    PROC Path_RobotLab(PERS wobjdata WO_Pastel)
        Path_vacio_ejecucion p_vacio_labSIR, 1, WO_Pastel, FALSE;
        index_vacio_destino:=25;
        Path_contacto_ejecucion p_contacto_labSIR, 1, 3, WO_Pastel, FALSE;
        Mover_en_contacto;
        TriggC p_contacto_labSIR{4},p_contacto_labSIR{5},Vel_Proceso,triggContactoCir,Z_Proceso,Prototipo_JSDaleman\WObj:=WO_Pastel;
        TriggL p_contacto_labSIR{6},Vel_Proceso,triggContacto,Z_Proceso,Prototipo_JSDaleman\WObj:=WO_Pastel;
        TriggC p_contacto_labSIR{7},p_contacto_labSIR{8},Vel_Proceso,triggContactoCir,Z_Proceso,Prototipo_JSDaleman\WObj:=WO_Pastel;
        Path_contacto_ejecucion p_contacto_labSIR, 9, 25, WO_Pastel, TRUE;
        Path_vacio_ejecucion p_vacio_labSIR, 2, WO_Pastel, FALSE;
        Path_contacto_ejecucion p_contacto_labSIR, 26, 94, WO_Pastel, TRUE;
        Path_vacio_ejecucion p_vacio_labSIR, 3, WO_Pastel, FALSE;
        Path_contacto_ejecucion p_contacto_labSIR, 95, 111, WO_Pastel, TRUE;
        Path_vacio_ejecucion p_vacio_labSIR, 4, WO_Pastel, FALSE;
        Path_contacto_ejecucion p_contacto_labSIR, 112, 125, WO_Pastel, TRUE;
        Path_vacio_ejecucion p_vacio_labSIR, 5, WO_Pastel, FALSE;
        index_vacio_destino:=131;
        Mover_a_contacto;
        TriggL p_contacto_labSIR{126},Vel_Acercamiento,triggContacto,Z_Acercamiento,Prototipo_JSDaleman\WObj:=WO_Pastel;
        Mover_en_contacto;
        TriggC p_contacto_labSIR{127},p_contacto_labSIR{128},Vel_Proceso,triggContactoCir,Z_Proceso,Prototipo_JSDaleman\WObj:=WO_Pastel;
        TriggC p_contacto_labSIR{129},p_contacto_labSIR{130},Vel_Proceso,triggContactoCir,Z_Proceso,Prototipo_JSDaleman\WObj:=WO_Pastel;
        Mover_a_vacio;
        TriggL p_contacto_labSIR{131},Vel_Acercamiento,triggContacto,Z_Acercamiento,Prototipo_JSDaleman\WObj:=WO_Pastel;
        Path_vacio_ejecucion p_vacio_labSIR, 6, WO_Pastel, FALSE;
        index_vacio_destino:=137;
        Mover_a_contacto;
        TriggL p_contacto_labSIR{132},Vel_Acercamiento,triggContacto,Z_Acercamiento,Prototipo_JSDaleman\WObj:=WO_Pastel;
        Mover_en_contacto;
        TriggC p_contacto_labSIR{133},p_contacto_labSIR{134},Vel_Proceso,triggContactoCir,Z_Proceso,Prototipo_JSDaleman\WObj:=WO_Pastel;
        TriggC p_contacto_labSIR{135},p_contacto_labSIR{136},Vel_Proceso,triggContactoCir,Z_Proceso,Prototipo_JSDaleman\WObj:=WO_Pastel;
        Mover_a_vacio;
        TriggL p_contacto_labSIR{137},Vel_Acercamiento,triggContacto,Z_Acercamiento,Prototipo_JSDaleman\WObj:=WO_Pastel;
        Path_vacio_ejecucion p_vacio_labSIR, 7, WO_Pastel, FALSE;
        index_vacio_destino:=143;
        Mover_a_contacto;
        TriggL p_contacto_labSIR{138},Vel_Acercamiento,triggContacto,Z_Acercamiento,Prototipo_JSDaleman\WObj:=WO_Pastel;
        Mover_en_contacto;
        TriggC p_contacto_labSIR{139},p_contacto_labSIR{140},Vel_Proceso,triggContactoCir,Z_Proceso,Prototipo_JSDaleman\WObj:=WO_Pastel;
        TriggC p_contacto_labSIR{141},p_contacto_labSIR{142},Vel_Proceso,triggContactoCir,Z_Proceso,Prototipo_JSDaleman\WObj:=WO_Pastel;
        Mover_a_vacio;
        TriggL p_contacto_labSIR{143},Vel_Acercamiento,triggContacto,Z_Acercamiento,Prototipo_JSDaleman\WObj:=WO_Pastel;
        Path_vacio_ejecucion p_vacio_labSIR, 8, WO_Pastel, FALSE;
        index_vacio_destino:=149;
        Mover_a_contacto;
        TriggL p_contacto_labSIR{144},Vel_Acercamiento,triggContacto,Z_Acercamiento,Prototipo_JSDaleman\WObj:=WO_Pastel;
        Mover_en_contacto;
        TriggC p_contacto_labSIR{145},p_contacto_labSIR{146},Vel_Proceso,triggContactoCir,Z_Proceso,Prototipo_JSDaleman\WObj:=WO_Pastel;
        TriggC p_contacto_labSIR{147},p_contacto_labSIR{148},Vel_Proceso,triggContactoCir,Z_Proceso,Prototipo_JSDaleman\WObj:=WO_Pastel;
        Mover_a_vacio;
        TriggL p_contacto_labSIR{149},Vel_Acercamiento,triggContacto,Z_Acercamiento,Prototipo_JSDaleman\WObj:=WO_Pastel;
        Path_vacio_ejecucion p_vacio_labSIR, 9, WO_Pastel, FALSE;
        index_vacio_destino:=155;
        Mover_a_contacto;
        TriggL p_contacto_labSIR{150},Vel_Acercamiento,triggContacto,Z_Acercamiento,Prototipo_JSDaleman\WObj:=WO_Pastel;
        Mover_en_contacto;
        TriggC p_contacto_labSIR{151},p_contacto_labSIR{152},Vel_Proceso,triggContactoCir,Z_Proceso,Prototipo_JSDaleman\WObj:=WO_Pastel;
        TriggC p_contacto_labSIR{153},p_contacto_labSIR{154},Vel_Proceso,triggContactoCir,Z_Proceso,Prototipo_JSDaleman\WObj:=WO_Pastel;
        Mover_a_vacio;
        TriggL p_contacto_labSIR{155},Vel_Acercamiento,triggContacto,Z_Acercamiento,Prototipo_JSDaleman\WObj:=WO_Pastel;
        Path_vacio_ejecucion p_vacio_labSIR, 10, WO_Pastel, FALSE;
        index_vacio_destino:=161;
        Mover_a_contacto;
        TriggL p_contacto_labSIR{156},Vel_Acercamiento,triggContacto,Z_Acercamiento,Prototipo_JSDaleman\WObj:=WO_Pastel;
        Mover_en_contacto;
        TriggC p_contacto_labSIR{157},p_contacto_labSIR{158},Vel_Proceso,triggContactoCir,Z_Proceso,Prototipo_JSDaleman\WObj:=WO_Pastel;
        TriggC p_contacto_labSIR{159},p_contacto_labSIR{160},Vel_Proceso,triggContactoCir,Z_Proceso,Prototipo_JSDaleman\WObj:=WO_Pastel;
        Mover_a_vacio;
        TriggL p_contacto_labSIR{161},Vel_Proceso,triggContacto,Z_Proceso,Prototipo_JSDaleman\WObj:=WO_Pastel;
    ENDPROC
    PROC Path_Tapa_LabSIR(PERS wobjdata WO_Pastel)
        Mover_en_vacio;
        MoveJ Target_Home_10,Vel_Vacio_Rap,Z_Vacio_Rap,Prototipo_JSDaleman\WObj:=wobj0;
        ReiniciarIndices;
        path_contacto_actual:="p_contacto_labSIR";
        path_vacio_actual:="p_vacio_labSIR";
        Path_RobotLab WO_Pastel;
        Path_LabSIR WO_Pastel;
        Mover_en_vacio;
        MoveJ Target_Home_10,Vel_Vacio_Rap,Z_Vacio_Rap,Prototipo_JSDaleman\WObj:=wobj0;
    ENDPROC
    PROC Path_LabSIR(PERS wobjdata WO_Pastel)
        Path_vacio_ejecucion p_vacio_labSIR, 11, WO_Pastel, FALSE;
        Path_contacto_ejecucion p_contacto_labSIR, 162, 170, WO_Pastel, TRUE;
        Path_vacio_ejecucion p_vacio_labSIR, 12, WO_Pastel, FALSE;
        Path_contacto_ejecucion p_contacto_labSIR, 171, 182, WO_Pastel, TRUE;
        Path_vacio_ejecucion p_vacio_labSIR, 13, WO_Pastel, FALSE;
        Path_contacto_ejecucion p_contacto_labSIR, 183, 188, WO_Pastel, TRUE;
        Path_vacio_ejecucion p_vacio_labSIR, 14, WO_Pastel, FALSE;
        Path_contacto_ejecucion p_contacto_labSIR, 189, 199, WO_Pastel, TRUE;
        Path_vacio_ejecucion p_vacio_labSIR, 15, WO_Pastel, FALSE;
        Path_contacto_ejecucion p_contacto_labSIR, 200, 205, WO_Pastel, TRUE;
        Path_vacio_ejecucion p_vacio_labSIR, 16, WO_Pastel, FALSE;
        Path_contacto_ejecucion p_contacto_labSIR, 206, 219, WO_Pastel, TRUE;
        Path_vacio_ejecucion p_vacio_labSIR, 17, WO_Pastel, FALSE;
        Path_contacto_ejecucion p_contacto_labSIR, 220, 226, WO_Pastel, TRUE;
        Path_vacio_ejecucion p_vacio_labSIR, 18, WO_Pastel, FALSE;
        Path_contacto_ejecucion p_contacto_labSIR, 227, 232, WO_Pastel, TRUE;
        Path_vacio_ejecucion p_vacio_labSIR, 19, WO_Pastel, FALSE;
        Path_contacto_ejecucion p_contacto_labSIR, 233, 256, WO_Pastel, TRUE;
    ENDPROC
    PROC Path_Frente_LabSIR(PERS wobjdata WO_Pastel)
        Mover_en_vacio;
        MoveJ Target_Home_10,Vel_Vacio_Rap,Z_Vacio_Rap,Prototipo_JSDaleman\WObj:=wobj0;
        MoveJ Target_Frente_10,Vel_Vacio,Z_VacioMov,Prototipo_JSDaleman\WObj:=WO_Pastel;
        MoveJ Target_Frente_20,Vel_Vacio,Z_VacioMov,Prototipo_JSDaleman\WObj:=WO_Pastel;
        ReiniciarIndices;
        path_contacto_actual:="p_contacto_labSIR_FrenteL";
        path_vacio_actual:="p_vacio_labSIR_FrenteL";
        Path_Chip WO_Pastel;
        Path_LetreroFrontal1_LabSIR WO_Pastel;
        Path_LetreroFrontal2_LabSIR WO_Pastel;
        Mover_en_vacio;
        MoveJ Target_Frente_20,Vel_Vacio,Z_VacioMov,Prototipo_JSDaleman\WObj:=WO_Pastel;
        MoveJ Target_Frente_10,Vel_Vacio,Z_VacioMov,Prototipo_JSDaleman\WObj:=WO_Pastel;
        MoveJ Target_Home_10,Vel_Vacio_Rap,Z_Vacio_Rap,Prototipo_JSDaleman\WObj:=wobj0;
        MoveJ Target_Frente_30,Vel_Vacio_Rap,Z_Vacio_Rap,Prototipo_JSDaleman\WObj:=WO_Pastel;
        MoveJ Target_Frente_40,Vel_Vacio_Rap,Z_Vacio_Rap,Prototipo_JSDaleman\WObj:=WO_Pastel;
        ReiniciarIndices;
        path_contacto_actual:="p_contacto_labSIR_FrenteR";
        path_vacio_actual:="p_vacio_labSIR_FrenteR";
        Path_Engranaje WO_Pastel;
        Path_LetreroFrontal3_LabSIR WO_Pastel;
        Path_LetreroFrontal4_LabSIR WO_Pastel;
        Mover_en_vacio;
        MoveJ Target_Frente_40,Vel_Vacio_Rap,Z_Vacio_Rap,Prototipo_JSDaleman\WObj:=WO_Pastel;
        MoveJ Target_Frente_30,Vel_Vacio_Rap,Z_Vacio_Rap,Prototipo_JSDaleman\WObj:=WO_Pastel;
        MoveJ Target_Home_10,Vel_Vacio_Rap,Z_Vacio_Rap,Prototipo_JSDaleman\WObj:=wobj0;
    ENDPROC
    PROC Path_Chip(PERS wobjdata WO_Pastel)
        Path_vacio_ejecucion p_vacio_labSIR_FrenteL, 1, WO_Pastel, FALSE;
        Path_contacto_ejecucion p_contacto_labSIR_FrenteL, 1, 50, WO_Pastel, TRUE;
        Path_vacio_ejecucion p_vacio_labSIR_FrenteL, 1, WO_Pastel, FALSE;
        Path_contacto_ejecucion p_contacto_labSIR_FrenteL, 51, 56, WO_Pastel, TRUE;
    ENDPROC
    PROC Path_LetreroFrontal1_LabSIR(PERS wobjdata WO_Pastel)
        Path_vacio_ejecucion p_vacio_labSIR_FrenteL, 3, WO_Pastel, FALSE;
        Path_contacto_ejecucion p_contacto_labSIR_FrenteL, 57, 60, WO_Pastel, TRUE;
        Path_vacio_ejecucion p_vacio_labSIR_FrenteL, 4, WO_Pastel, FALSE;
        Path_contacto_ejecucion p_contacto_labSIR_FrenteL, 61, 74, WO_Pastel, TRUE;
        Path_vacio_ejecucion p_vacio_labSIR_FrenteL, 5, WO_Pastel, FALSE;
        Path_contacto_ejecucion p_contacto_labSIR_FrenteL, 75, 92, WO_Pastel, TRUE;
        Path_vacio_ejecucion p_vacio_labSIR_FrenteL, 6, WO_Pastel, FALSE;
        Path_contacto_ejecucion p_contacto_labSIR_FrenteL, 93, 116, WO_Pastel, TRUE;
        Path_vacio_ejecucion p_vacio_labSIR_FrenteL, 7, WO_Pastel, FALSE;
        Path_contacto_ejecucion p_contacto_labSIR_FrenteL, 117, 122, WO_Pastel, TRUE;
        Path_vacio_ejecucion p_vacio_labSIR_FrenteL, 8, WO_Pastel, FALSE;
        Path_contacto_ejecucion p_contacto_labSIR_FrenteL, 123, 140, WO_Pastel, TRUE;
        Path_vacio_ejecucion p_vacio_labSIR_FrenteL, 9, WO_Pastel, FALSE;
        Path_contacto_ejecucion p_contacto_labSIR_FrenteL, 141, 149, WO_Pastel, TRUE;
        Path_vacio_ejecucion p_vacio_labSIR_FrenteL, 10, WO_Pastel, FALSE;
        Path_contacto_ejecucion p_contacto_labSIR_FrenteL, 150, 174, WO_Pastel, TRUE;
        Path_vacio_ejecucion p_vacio_labSIR_FrenteL, 11, WO_Pastel, FALSE;
        Path_contacto_ejecucion p_contacto_labSIR_FrenteL, 175, 183, WO_Pastel, TRUE;
        Path_vacio_ejecucion p_vacio_labSIR_FrenteL, 12, WO_Pastel, FALSE;
        Path_contacto_ejecucion p_contacto_labSIR_FrenteL, 184, 186, WO_Pastel, TRUE;
        Path_vacio_ejecucion p_vacio_labSIR_FrenteL, 13, WO_Pastel, FALSE;
        index_vacio_destino:=188;
        Mover_a_contacto;
        TriggL p_contacto_labSIR_FrenteL{187},Vel_Acercamiento,triggContacto,Z_Acercamiento,Prototipo_JSDaleman\WObj:=WO_Pastel;
        Mover_en_contacto;
        TriggL p_contacto_labSIR_FrenteL{188},Vel_Acercamiento_Lateral,triggContacto,Z_Acercamiento,Prototipo_JSDaleman\WObj:=WO_Pastel;
        Path_vacio_ejecucion p_vacio_labSIR_FrenteL, 14, WO_Pastel, FALSE;
        Path_contacto_ejecucion p_contacto_labSIR_FrenteL, 189, 212, WO_Pastel, TRUE;
    ENDPROC
    PROC Path_LetreroFrontal2_LabSIR(PERS wobjdata WO_Pastel)
        Path_vacio_ejecucion p_vacio_labSIR_FrenteL, 15, WO_Pastel, FALSE;
        Path_contacto_ejecucion p_contacto_labSIR_FrenteL, 213, 238, WO_Pastel, TRUE;
        Path_vacio_ejecucion p_vacio_labSIR_FrenteL, 16, WO_Pastel, FALSE;
        Path_contacto_ejecucion p_contacto_labSIR_FrenteL, 239, 262, WO_Pastel, TRUE;
        Path_vacio_ejecucion p_vacio_labSIR_FrenteL, 17, WO_Pastel, FALSE;
        Path_contacto_ejecucion p_contacto_labSIR_FrenteL, 263, 273, WO_Pastel, TRUE;
        Path_vacio_ejecucion p_vacio_labSIR_FrenteL, 18, WO_Pastel, FALSE;
        Path_contacto_ejecucion p_contacto_labSIR_FrenteL, 274, 287, WO_Pastel, TRUE;
        Path_vacio_ejecucion p_vacio_labSIR_FrenteL, 19, WO_Pastel, FALSE;
        Path_contacto_ejecucion p_contacto_labSIR_FrenteL, 288, 307, WO_Pastel, TRUE;
        Path_vacio_ejecucion p_vacio_labSIR_FrenteL, 20, WO_Pastel, FALSE;
        Path_contacto_ejecucion p_contacto_labSIR_FrenteL, 308, 341, WO_Pastel, TRUE;
        Path_vacio_ejecucion p_vacio_labSIR_FrenteL, 21, WO_Pastel, FALSE;
        Path_contacto_ejecucion p_contacto_labSIR_FrenteL, 342, 344, WO_Pastel, TRUE;
        Path_vacio_ejecucion p_vacio_labSIR_FrenteL, 22, WO_Pastel, FALSE;
        Path_contacto_ejecucion p_contacto_labSIR_FrenteL, 345, 346, WO_Pastel, TRUE;
        Path_vacio_ejecucion p_vacio_labSIR_FrenteL, 23, WO_Pastel, FALSE;
        Path_contacto_ejecucion p_contacto_labSIR_FrenteL, 347, 350, WO_Pastel, TRUE;
        Path_vacio_ejecucion p_vacio_labSIR_FrenteL, 24, WO_Pastel, FALSE;
        Path_contacto_ejecucion p_contacto_labSIR_FrenteL, 351, 370, WO_Pastel, TRUE;
        Path_vacio_ejecucion p_vacio_labSIR_FrenteL, 25, WO_Pastel, FALSE;
        Path_contacto_ejecucion p_contacto_labSIR_FrenteL, 371, 379, WO_Pastel, TRUE;
        Path_vacio_ejecucion p_vacio_labSIR_FrenteL, 26, WO_Pastel, FALSE;
        Path_contacto_ejecucion p_contacto_labSIR_FrenteL, 380, 391, WO_Pastel, TRUE;
        Path_vacio_ejecucion p_vacio_labSIR_FrenteL, 27, WO_Pastel, FALSE;
        Path_contacto_ejecucion p_contacto_labSIR_FrenteL, 392, 394, WO_Pastel, TRUE;
    ENDPROC
    PROC Path_Engranaje(PERS wobjdata WO_Pastel)
        Path_vacio_ejecucion p_vacio_labSIR_FrenteR, 1, WO_Pastel, FALSE;
        Path_contacto_ejecucion p_contacto_labSIR_FrenteR, 1, 78, WO_Pastel, TRUE;
        Path_vacio_ejecucion p_vacio_labSIR_FrenteR, 2, WO_Pastel, FALSE;
        Path_contacto_ejecucion p_contacto_labSIR_FrenteR, 79, 97, WO_Pastel, TRUE;
    ENDPROC
    PROC Path_LetreroFrontal3_LabSIR(PERS wobjdata WO_Pastel)
        Path_vacio_ejecucion p_vacio_labSIR_FrenteR, 3, WO_Pastel, FALSE;
        Path_contacto_ejecucion p_contacto_labSIR_FrenteR, 98, 121, WO_Pastel, TRUE;
        Path_vacio_ejecucion p_vacio_labSIR_FrenteR, 4, WO_Pastel, FALSE;
        Path_contacto_ejecucion p_contacto_labSIR_FrenteR, 122, 150, WO_Pastel, TRUE;
        Path_vacio_ejecucion p_vacio_labSIR_FrenteR, 5, WO_Pastel, FALSE;
        Path_contacto_ejecucion p_contacto_labSIR_FrenteR, 151, 163, WO_Pastel, TRUE;
        Path_vacio_ejecucion p_vacio_labSIR_FrenteR, 6, WO_Pastel, FALSE;
        Path_contacto_ejecucion p_contacto_labSIR_FrenteR, 164, 187, WO_Pastel, TRUE;
        Path_vacio_ejecucion p_vacio_labSIR_FrenteR, 7, WO_Pastel, FALSE;
        Path_contacto_ejecucion p_contacto_labSIR_FrenteR, 188, 198, WO_Pastel, TRUE;
        Path_vacio_ejecucion p_vacio_labSIR_FrenteR, 8, WO_Pastel, FALSE;
        Path_contacto_ejecucion p_contacto_labSIR_FrenteR, 199, 218, WO_Pastel, TRUE;
        Path_vacio_ejecucion p_vacio_labSIR_FrenteR, 9, WO_Pastel, FALSE;
        Path_contacto_ejecucion p_contacto_labSIR_FrenteR, 219, 221, WO_Pastel, TRUE;
        Path_vacio_ejecucion p_vacio_labSIR_FrenteR, 10, WO_Pastel, FALSE;
        Path_contacto_ejecucion p_contacto_labSIR_FrenteR, 222, 223, WO_Pastel, TRUE;
        Path_vacio_ejecucion p_vacio_labSIR_FrenteR, 11, WO_Pastel, FALSE;
        Path_contacto_ejecucion p_contacto_labSIR_FrenteR, 224, 242, WO_Pastel, TRUE;
        Path_vacio_ejecucion p_vacio_labSIR_FrenteR, 12, WO_Pastel, FALSE;
        Path_contacto_ejecucion p_contacto_labSIR_FrenteR, 243, 264, WO_Pastel, TRUE;
        Path_vacio_ejecucion p_vacio_labSIR_FrenteR, 13, WO_Pastel, FALSE;
        Path_contacto_ejecucion p_contacto_labSIR_FrenteR, 265, 281, WO_Pastel, TRUE;
    ENDPROC
    PROC Path_LetreroFrontal4_LabSIR(PERS wobjdata WO_Pastel)
        Path_vacio_ejecucion p_vacio_labSIR_FrenteR, 14, WO_Pastel, FALSE;
        Path_contacto_ejecucion p_contacto_labSIR_FrenteR, 282, 293, WO_Pastel, TRUE;
        Path_vacio_ejecucion p_vacio_labSIR_FrenteR, 15, WO_Pastel, FALSE;
        Path_contacto_ejecucion p_contacto_labSIR_FrenteR, 294, 317, WO_Pastel, TRUE;
        Path_vacio_ejecucion p_vacio_labSIR_FrenteR, 16, WO_Pastel, FALSE;
        Path_contacto_ejecucion p_contacto_labSIR_FrenteR, 318, 332, WO_Pastel, TRUE;
        Path_vacio_ejecucion p_vacio_labSIR_FrenteR, 17, WO_Pastel, FALSE;
        Path_contacto_ejecucion p_contacto_labSIR_FrenteR, 333, 350, WO_Pastel, TRUE;
        Path_vacio_ejecucion p_vacio_labSIR_FrenteR, 18, WO_Pastel, FALSE;
        Path_contacto_ejecucion p_contacto_labSIR_FrenteR, 351, 360, WO_Pastel, TRUE;
        Path_vacio_ejecucion p_vacio_labSIR_FrenteR, 19, WO_Pastel, FALSE;
        Path_contacto_ejecucion p_contacto_labSIR_FrenteR, 361, 363, WO_Pastel, TRUE;
        Path_vacio_ejecucion p_vacio_labSIR_FrenteR, 20, WO_Pastel, FALSE;
        Path_contacto_ejecucion p_contacto_labSIR_FrenteR, 364, 365, WO_Pastel, TRUE;
        Path_vacio_ejecucion p_vacio_labSIR_FrenteR, 21, WO_Pastel, FALSE;
        Path_contacto_ejecucion p_contacto_labSIR_FrenteR, 366, 370, WO_Pastel, TRUE;
        Path_vacio_ejecucion p_vacio_labSIR_FrenteR, 22, WO_Pastel, FALSE;
        Path_contacto_ejecucion p_contacto_labSIR_FrenteR, 371, 394, WO_Pastel, TRUE;
        Path_vacio_ejecucion p_vacio_labSIR_FrenteR, 23, WO_Pastel, FALSE;
        Path_contacto_ejecucion p_contacto_labSIR_FrenteR, 395, 410, WO_Pastel, TRUE;
        Path_vacio_ejecucion p_vacio_labSIR_FrenteR, 24, WO_Pastel, FALSE;
        Path_contacto_ejecucion p_contacto_labSIR_FrenteR, 411, 430, WO_Pastel, TRUE;
        Path_vacio_ejecucion p_vacio_labSIR_FrenteR, 25, WO_Pastel, FALSE;
        Path_contacto_ejecucion p_contacto_labSIR_FrenteR, 431, 448, WO_Pastel, TRUE;
    ENDPROC
ENDMODULE

--- Controller Data/IRB140_LabSIR/RAPID/TASK1/PROGMOD/Mecatronica25.mod ---
MODULE Mecatronica25
    !***********************************************************
    !
    ! Modulo:  Mecatronica25
    !
    ! Descripci?n:
    !   Modulo con rutinas para decoracion con el motivo 25 a?os de ingeneria mecatronica
    !
    ! Autor: Juan_Daleman
    !
    ! Versi?n: 1.0
    !
    !***********************************************************

    CONST robtarget Target_Tap25_10:=[[71.235002268,-92.346037462,-20.000000611],[0.707106779,-0.000000013,0.00000001,0.707106783],[-1,0,-1,0],[9E+09,9E+09,9E+09,9E+09,9E+09,9E+09]];
    CONST robtarget Target_Tap25_20:=[[71.235,-92.346,-2.358],[0.707106781,0,0,0.707106781],[0,0,0,0],[9E+09,9E+09,9E+09,9E+09,9E+09,9E+09]];
    CONST robtarget Target_Tap25_30:=[[70.898,-75.837,-2.361],[0.707106781,0,0,0.707106781],[0,0,0,0],[9E+09,9E+09,9E+09,9E+09,9E+09,9E+09]];
    CONST robtarget Target_Tap25_40:=[[63.811,-92.424,-2.425],[0.707106781,0,0,0.707106781],[0,0,0,0],[9E+09,9E+09,9E+09,9E+09,9E+09,9E+09]];
    CONST robtarget Target_Tap25_50:=[[56.589,-76.018,-2.491],[0.707106781,0,0,0.707106781],[0,0,0,0],[9E+09,9E+09,9E+09,9E+09,9E+09,9E+09]];
    CONST robtarget Target_Tap25_60:=[[56.589,-92.474,-2.491],[0.707106781,0,0,0.707106781],[0,0,0,0],[9E+09,9E+09,9E+09,9E+09,9E+09,9E+09]];
    CONST robtarget Target_Tap25_70:=[[56.589,-92.474,-20],[0.707106781,0,0,0.707106781],[0,0,0,0],[9E+09,9E+09,9E+09,9E+09,9E+09,9E+09]];
    CONST robtarget Target_Tap25_80:=[[41.198,-88.513,-20],[0.707106781,0,0,0.707106781],[0,0,0,0],[9E+09,9E+09,9E+09,9E+09,9E+09,9E+09]];
    CONST robtarget Target_Tap25_90:=[[41.18,-88.446,-2.63],[0.707106781,0,0,0.707106781],[0,0,0,0],[9E+09,9E+09,9E+09,9E+09,9E+09,9E+09]];
    CONST robtarget Target_Tap25_100:=[[47.311,-92.769,-2.575],[0.707106781,0,0,0.707106781],[0,0,0,0],[9E+09,9E+09,9E+09,9E+09,9E+09,9E+09]];
    CONST robtarget Target_Tap25_110:=[[53.192,-86.979,-2.521],[0.707106781,0,0,0.707106781],[0,0,0,0],[9E+09,9E+09,9E+09,9E+09,9E+09,9E+09]];
    CONST robtarget Target_Tap25_120:=[[47.79,-79.621,-2.57],[0.707106781,0,0,0.707106781],[0,0,0,0],[9E+09,9E+09,9E+09,9E+09,9E+09,9E+09]];
    CONST robtarget Target_Tap25_130:=[[40.922,-86.876,-2.633],[0.707106781,0,0,0.707106781],[-1,0,-2,0],[9E+09,9E+09,9E+09,9E+09,9E+09,9E+09]];
    CONST robtarget Target_Tap25_140:=[[49.328,-87.108,-2.556],[0.707106781,0,0,0.707106781],[0,0,0,0],[9E+09,9E+09,9E+09,9E+09,9E+09,9E+09]];
    CONST robtarget Target_Tap25_150:=[[49.328,-87.108,-20],[0.707106781,0,0,0.707106781],[0,0,0,0],[9E+09,9E+09,9E+09,9E+09,9E+09,9E+09]];
    CONST robtarget Target_Tap25_160:=[[27.912,-88.405,-19.751],[0.707106781,0,0,0.707106781],[-1,0,-1,0],[9E+09,9E+09,9E+09,9E+09,9E+09,9E+09]];
    CONST robtarget Target_Tap25_170:=[[27.863,-88.19,-2.751],[0.707106781,0,0,0.707106781],[0,0,0,0],[9E+09,9E+09,9E+09,9E+09,9E+09,9E+09]];
    CONST robtarget Target_Tap25_180:=[[35.24,-92.83,-2.684],[0.707106781,0,0,0.707106781],[0,0,0,0],[9E+09,9E+09,9E+09,9E+09,9E+09,9E+09]];
    CONST robtarget Target_Tap25_190:=[[39.889,-85.357,-2.642],[0.707106781,0,0,0.707106781],[0,0,0,0],[9E+09,9E+09,9E+09,9E+09,9E+09,9E+09]];
    CONST robtarget Target_Tap25_200:=[[33.589,-79.684,-2.699],[0.707106781,0,0,0.707106781],[0,0,0,0],[9E+09,9E+09,9E+09,9E+09,9E+09,9E+09]];
    CONST robtarget Target_Tap25_210:=[[27.903,-84.371,-2.751],[0.707106781,0,0,0.707106781],[0,0,0,0],[9E+09,9E+09,9E+09,9E+09,9E+09,9E+09]];
    CONST robtarget Target_Tap25_220:=[[27.903,-84.371,-19.751],[0.707106781,0,0,0.707106781],[0,0,0,0],[9E+09,9E+09,9E+09,9E+09,9E+09,9E+09]];
    CONST robtarget Target_Tap25_230:=[[15.792,-80.111,-20],[0.707106781,0,0,0.707106781],[0,0,0,0],[9E+09,9E+09,9E+09,9E+09,9E+09,9E+09]];
    CONST robtarget Target_Tap25_240:=[[15.792,-80.111,-2.861],[0.707106781,0,0,0.707106781],[0,0,0,0],[9E+09,9E+09,9E+09,9E+09,9E+09,9E+09]];
    CONST robtarget Target_Tap25_250:=[[15.593,-92.922,-2.863],[0.707106781,0,0,0.707106781],[0,0,0,0],[9E+09,9E+09,9E+09,9E+09,9E+09,9E+09]];
    CONST robtarget Target_Tap25_260:=[[17.701,-91.357,-2.843],[0.707106781,0,0,0.707106781],[0,0,0,0],[9E+09,9E+09,9E+09,9E+09,9E+09,9E+09]];
    CONST robtarget Target_Tap25_270:=[[22.44,-93.01,-2.8],[0.707106781,0,0,0.707106781],[0,0,0,0],[9E+09,9E+09,9E+09,9E+09,9E+09,9E+09]];
    CONST robtarget Target_Tap25_280:=[[26.795,-87.318,-2.761],[0.707106781,0,0,0.707106781],[0,0,0,0],[9E+09,9E+09,9E+09,9E+09,9E+09,9E+09]];
    CONST robtarget Target_Tap25_290:=[[25.214,-81.575,-2.775],[0.707106781,0,0,0.707106781],[0,0,0,0],[9E+09,9E+09,9E+09,9E+09,9E+09,9E+09]];
    CONST robtarget Target_Tap25_300:=[[21.612,-79.848,-2.808],[0.707106781,0,0,0.707106781],[0,0,0,0],[9E+09,9E+09,9E+09,9E+09,9E+09,9E+09]];
    CONST robtarget Target_Tap25_310:=[[17.639,-81.422,-2.844],[0.707106781,0,0,0.707106781],[0,0,0,0],[9E+09,9E+09,9E+09,9E+09,9E+09,9E+09]];
    CONST robtarget Target_Tap25_320:=[[17.639,-81.422,-20],[0.707106781,0,0,0.707106781],[0,0,0,0],[9E+09,9E+09,9E+09,9E+09,9E+09,9E+09]];
    CONST robtarget Target_Tap25_330:=[[9.176,-76.919,-20],[0.707106781,0,0,0.707106781],[0,0,0,0],[9E+09,9E+09,9E+09,9E+09,9E+09,9E+09]];
    CONST robtarget Target_Tap25_340:=[[9.176,-76.919,-2.921],[0.707106781,0,0,0.707106781],[0,0,0,0],[9E+09,9E+09,9E+09,9E+09,9E+09,9E+09]];
    CONST robtarget Target_Tap25_350:=[[10.914,-80.118,-2.905],[0.707106781,0,0,0.707106781],[0,0,0,0],[9E+09,9E+09,9E+09,9E+09,9E+09,9E+09]];
    CONST robtarget Target_Tap25_360:=[[12.324,-80.117,-2.892],[0.707106781,0,0,0.707106781],[0,0,0,0],[9E+09,9E+09,9E+09,9E+09,9E+09,9E+09]];
    CONST robtarget Target_Tap25_370:=[[4.821,-80.264,-2.96],[0.707106781,0,0,0.707106781],[0,0,0,0],[9E+09,9E+09,9E+09,9E+09,9E+09,9E+09]];
    CONST robtarget Target_Tap25_380:=[[6.952,-80.063,-2.941],[0.707106781,0,0,0.707106781],[0,0,0,0],[9E+09,9E+09,9E+09,9E+09,9E+09,9E+09]];
    CONST robtarget Target_Tap25_390:=[[9.179,-76.919,-2.921],[0.707106781,0,0,0.707106781],[0,0,0,0],[9E+09,9E+09,9E+09,9E+09,9E+09,9E+09]];
    CONST robtarget Target_Tap25_400:=[[8.458,-92.812,-2.927],[0.707106781,0,0,0.707106781],[0,0,0,0],[9E+09,9E+09,9E+09,9E+09,9E+09,9E+09]];
    CONST robtarget Target_Tap25_410:=[[4.611,-93.079,-2.962],[0.707106781,0,0,0.707106781],[0,0,0,0],[9E+09,9E+09,9E+09,9E+09,9E+09,9E+09]];
    CONST robtarget Target_Tap25_420:=[[4.611,-93.079,-20],[0.707106781,0,0,0.707106781],[0,0,0,0],[9E+09,9E+09,9E+09,9E+09,9E+09,9E+09]];
    CONST robtarget Target_Tap25_430:=[[0.994,-93.119,-20],[0.707106781,0,0,0.707106781],[0,0,0,0],[9E+09,9E+09,9E+09,9E+09,9E+09,9E+09]];
    CONST robtarget Target_Tap25_440:=[[0.972,-93.119,-2.995],[0.707106781,0,0,0.707106781],[0,0,0,0],[9E+09,9E+09,9E+09,9E+09,9E+09,9E+09]];
    CONST robtarget Target_Tap25_450:=[[1.504,-80.221,-2.99],[0.707106781,0,0,0.707106781],[0,0,0,0],[9E+09,9E+09,9E+09,9E+09,9E+09,9E+09]];
    CONST robtarget Target_Tap25_460:=[[-1.051,-82.034,-3.014],[0.707106781,0,0,0.707106781],[0,0,0,0],[9E+09,9E+09,9E+09,9E+09,9E+09,9E+09]];
    CONST robtarget Target_Tap25_470:=[[-4.392,-80.165,-3.044],[0.707106781,0,0,0.707106781],[0,0,0,0],[9E+09,9E+09,9E+09,9E+09,9E+09,9E+09]];
    CONST robtarget Target_Tap25_480:=[[-4.392,-80.165,-20],[0.707106781,0,0,0.707106781],[0,0,0,0],[9E+09,9E+09,9E+09,9E+09,9E+09,9E+09]];
    CONST robtarget Target_Tap25_490:=[[-9.253,-77.852,-20],[0.707106781,0,0,0.707106781],[0,0,0,0],[9E+09,9E+09,9E+09,9E+09,9E+09,9E+09]];
    CONST robtarget Target_Tap25_500:=[[-9.253,-77.852,-3.088],[0.707106781,0,0,0.707106781],[0,0,0,0],[9E+09,9E+09,9E+09,9E+09,9E+09,9E+09]];
    CONST robtarget Target_Tap25_510:=[[-14.717,-75.57,-3.138],[0.707106781,0,0,0.707106781],[0,0,0,0],[9E+09,9E+09,9E+09,9E+09,9E+09,9E+09]];
    CONST robtarget Target_Tap25_520:=[[-14.718,-75.491,-20],[0.707106781,0,0,0.707106781],[0,0,0,0],[9E+09,9E+09,9E+09,9E+09,9E+09,9E+09]];
    CONST robtarget Target_Tap25_530:=[[-11.341,-80.235,-20],[0.707106781,0,0,0.707106781],[0,0,0,0],[9E+09,9E+09,9E+09,9E+09,9E+09,9E+09]];
    CONST robtarget Target_Tap25_540:=[[-11.341,-80.235,-3.107],[0.707106781,0,0,0.707106781],[0,0,0,0],[9E+09,9E+09,9E+09,9E+09,9E+09,9E+09]];
    CONST robtarget Target_Tap25_550:=[[-18.028,-85.783,-3.168],[0.707106781,0,0,0.707106781],[0,0,0,0],[9E+09,9E+09,9E+09,9E+09,9E+09,9E+09]];
    CONST robtarget Target_Tap25_560:=[[-10.892,-93.389,-3.103],[0.707106781,0,0,0.707106781],[0,0,0,0],[9E+09,9E+09,9E+09,9E+09,9E+09,9E+09]];
    CONST robtarget Target_Tap25_570:=[[-5.378,-85.572,-3.053],[0.707106781,0,0,0.707106781],[0,0,0,0],[9E+09,9E+09,9E+09,9E+09,9E+09,9E+09]];
    CONST robtarget Target_Tap25_580:=[[-11.36,-80.236,-3.107],[0.707106781,0,0,0.707106781],[0,0,0,0],[9E+09,9E+09,9E+09,9E+09,9E+09,9E+09]];
    CONST robtarget Target_Tap25_590:=[[-11.36,-80.236,-20],[0.707106781,0,0,0.707106781],[0,0,0,0],[9E+09,9E+09,9E+09,9E+09,9E+09,9E+09]];
    CONST robtarget Target_Tap25_600:=[[-21.618,-93.367,-20],[0.707106781,0,0,0.707106781],[0,0,0,0],[9E+09,9E+09,9E+09,9E+09,9E+09,9E+09]];
    CONST robtarget Target_Tap25_610:=[[-21.618,-93.367,-3.2],[0.707106781,0,0,0.707106781],[0,0,0,0],[9E+09,9E+09,9E+09,9E+09,9E+09,9E+09]];
    CONST robtarget Target_Tap25_620:=[[-21.187,-80.498,-3.196],[0.707106781,0,0,0.707106781],[0,0,0,0],[9E+09,9E+09,9E+09,9E+09,9E+09,9E+09]];
    CONST robtarget Target_Tap25_630:=[[-23.739,-81.876,-3.22],[0.707106781,0,0,0.707106781],[0,0,0,0],[9E+09,9E+09,9E+09,9E+09,9E+09,9E+09]];
    CONST robtarget Target_Tap25_640:=[[-28.5,-80.587,-3.263],[0.707106781,0,0,0.707106781],[0,0,0,0],[9E+09,9E+09,9E+09,9E+09,9E+09,9E+09]];
    CONST robtarget Target_Tap25_650:=[[-31.948,-84.819,-3.294],[0.707106781,0,0,0.707106781],[0,0,0,0],[9E+09,9E+09,9E+09,9E+09,9E+09,9E+09]];
    CONST robtarget Target_Tap25_660:=[[-31.767,-93.351,-3.292],[0.707106781,0,0,0.707106781],[0,0,0,0],[9E+09,9E+09,9E+09,9E+09,9E+09,9E+09]];
    CONST robtarget Target_Tap25_670:=[[-31.767,-93.351,-20],[0.707106781,0,0,0.707106781],[0,0,0,0],[9E+09,9E+09,9E+09,9E+09,9E+09,9E+09]];
    CONST robtarget Target_Tap25_680:=[[-35.856,-93.259,-20],[0.707106781,0,0,0.707106781],[0,0,0,0],[9E+09,9E+09,9E+09,9E+09,9E+09,9E+09]];
    CONST robtarget Target_Tap25_690:=[[-35.856,-93.259,-3.33],[0.707106781,0,0,0.707106781],[0,0,0,0],[9E+09,9E+09,9E+09,9E+09,9E+09,9E+09]];
    CONST robtarget Target_Tap25_700:=[[-36.105,-80.635,-3.332],[0.707106781,0,0,0.707106781],[0,0,0,0],[9E+09,9E+09,9E+09,9E+09,9E+09,9E+09]];
    CONST robtarget Target_Tap25_710:=[[-36.105,-80.635,-20],[0.707106781,0,0,0.707106781],[0,0,0,0],[9E+09,9E+09,9E+09,9E+09,9E+09,9E+09]];
    CONST robtarget Target_Tap25_720:=[[-36.199,-75.007,-20],[0.707106781,0,0,0.707106781],[0,0,0,0],[9E+09,9E+09,9E+09,9E+09,9E+09,9E+09]];
    CONST robtarget Target_Tap25_730:=[[-36.199,-75.007,-0.333],[0.707106781,0,0,0.707106781],[0,0,0,0],[9E+09,9E+09,9E+09,9E+09,9E+09,9E+09]];
    CONST robtarget Target_Tap25_740:=[[-36.286,-75.017,-20],[0.707106781,0,0,0.707106781],[0,0,0,0],[9E+09,9E+09,9E+09,9E+09,9E+09,9E+09]];
    CONST robtarget Target_Tap25_750:=[[-51.57,-89.064,-20],[0.707106781,0,0,0.707106781],[0,0,0,0],[9E+09,9E+09,9E+09,9E+09,9E+09,9E+09]];
    CONST robtarget Target_Tap25_760:=[[-51.674,-89.141,-3.473],[0.707106781,0,0,0.707106781],[0,0,0,0],[9E+09,9E+09,9E+09,9E+09,9E+09,9E+09]];
    CONST robtarget Target_Tap25_770:=[[-45.29,-93.794,-3.415],[0.707106781,0,0,0.707106781],[0,0,0,0],[9E+09,9E+09,9E+09,9E+09,9E+09,9E+09]];
    CONST robtarget Target_Tap25_780:=[[-39.461,-87.342,-3.362],[0.707106781,0,0,0.707106781],[0,0,0,0],[9E+09,9E+09,9E+09,9E+09,9E+09,9E+09]];
    CONST robtarget Target_Tap25_790:=[[-44.602,-80.683,-3.409],[0.707106781,0,0,0.707106781],[0,0,0,0],[9E+09,9E+09,9E+09,9E+09,9E+09,9E+09]];
    CONST robtarget Target_Tap25_800:=[[-51.56,-85.266,-3.472],[0.707106781,0,0,0.707106781],[0,0,0,0],[9E+09,9E+09,9E+09,9E+09,9E+09,9E+09]];
    CONST robtarget Target_Tap25_810:=[[-51.56,-85.266,-20],[0.707106781,0,0,0.707106781],[0,0,0,0],[9E+09,9E+09,9E+09,9E+09,9E+09,9E+09]];
    CONST robtarget Target_Tap25_820:=[[-63.731,-80.974,-20],[0.707106781,0,0,0.707106781],[0,0,0,0],[9E+09,9E+09,9E+09,9E+09,9E+09,9E+09]];
    CONST robtarget Target_Tap25_830:=[[-63.75,-80.975,-3.583],[0.707106781,0,0,0.707106781],[0,0,0,0],[9E+09,9E+09,9E+09,9E+09,9E+09,9E+09]];
    CONST robtarget Target_Tap25_840:=[[-63.89,-93.832,-3.584],[0.707106781,0,0,0.707106781],[0,0,0,0],[9E+09,9E+09,9E+09,9E+09,9E+09,9E+09]];
    CONST robtarget Target_Tap25_850:=[[-61.748,-92.459,-3.565],[0.707106781,0,0,0.707106781],[0,0,0,0],[9E+09,9E+09,9E+09,9E+09,9E+09,9E+09]];
    CONST robtarget Target_Tap25_860:=[[-56.209,-93.673,-3.514],[0.707106781,0,0,0.707106781],[0,0,0,0],[9E+09,9E+09,9E+09,9E+09,9E+09,9E+09]];
    CONST robtarget Target_Tap25_870:=[[-52.803,-85.856,-3.483],[0.707106781,0,0,0.707106781],[0,0,0,0],[9E+09,9E+09,9E+09,9E+09,9E+09,9E+09]];
    CONST robtarget Target_Tap25_880:=[[-56.502,-80.983,-3.517],[0.707106781,0,0,0.707106781],[0,0,0,0],[9E+09,9E+09,9E+09,9E+09,9E+09,9E+09]];
    CONST robtarget Target_Tap25_890:=[[-61.855,-82.29,-3.566],[0.707106781,0,0,0.707106781],[0,0,0,0],[9E+09,9E+09,9E+09,9E+09,9E+09,9E+09]];
    CONST robtarget Target_Tap25_900:=[[-61.855,-82.29,-20],[0.707106781,0,0,0.707106781],[0,0,0,0],[9E+09,9E+09,9E+09,9E+09,9E+09,9E+09]];
    CONST robtarget Target_Tap25_910:=[[5.931,-29.884,-20],[0.707106781,0,0,0.707106781],[0,0,0,0],[9E+09,9E+09,9E+09,9E+09,9E+09,9E+09]];
    CONST robtarget Target_Tap25_920:=[[5.931,-29.884,-1.95],[0.707106781,0,0,0.707106781],[0,0,0,0],[9E+09,9E+09,9E+09,9E+09,9E+09,9E+09]];
    CONST robtarget Target_Tap25_930:=[[-28.804,-64.72,-2.266],[0.707106781,0,0,0.707106781],[0,0,0,0],[9E+09,9E+09,9E+09,9E+09,9E+09,9E+09]];
    CONST robtarget Target_Tap25_940:=[[-64.967,-28.761,-2.594],[0.707106781,0,0,0.707106781],[0,0,0,0],[9E+09,9E+09,9E+09,9E+09,9E+09,9E+09]];
    CONST robtarget Target_Tap25_950:=[[-48.605,2.796,-2.445],[0.707106781,0,0,0.707106781],[0,0,0,0],[9E+09,9E+09,9E+09,9E+09,9E+09,9E+09]];
    CONST robtarget Target_Tap25_960:=[[-31.151,8.724,-2.287],[0.707106781,0,0,0.707106781],[0,0,0,0],[9E+09,9E+09,9E+09,9E+09,9E+09,9E+09]];
    CONST robtarget Target_Tap25_970:=[[-15.41,9.23,-2.144],[0.707106781,0,0,0.707106781],[0,0,0,0],[9E+09,9E+09,9E+09,9E+09,9E+09,9E+09]];
    CONST robtarget Target_Tap25_980:=[[-15.51,26.958,-2.145],[0.707106781,0,0,0.707106781],[0,0,0,0],[9E+09,9E+09,9E+09,9E+09,9E+09,9E+09]];
    CONST robtarget Target_Tap25_990:=[[-57.918,26.492,-2.53],[0.707106781,0,0,0.707106781],[0,0,0,0],[9E+09,9E+09,9E+09,9E+09,9E+09,9E+09]];
    CONST robtarget Target_Tap25_1000:=[[-57.918,26.492,-20],[0.707106781,0,0,0.707106781],[0,0,0,0],[9E+09,9E+09,9E+09,9E+09,9E+09,9E+09]];
    CONST robtarget Target_Tap25_1010:=[[-58.237,44.312,-20],[0.707106781,0,0,0.707106781],[0,0,0,0],[9E+09,9E+09,9E+09,9E+09,9E+09,9E+09]];
    CONST robtarget Target_Tap25_1020:=[[-58.218,44.658,-2.533],[0.707106781,0,0,0.707106781],[0,0,0,0],[9E+09,9E+09,9E+09,9E+09,9E+09,9E+09]];
    CONST robtarget Target_Tap25_1030:=[[2.688,45.238,-1.98],[0.707106781,0,0,0.707106781],[0,0,0,0],[9E+09,9E+09,9E+09,9E+09,9E+09,9E+09]];
    CONST robtarget Target_Tap25_1040:=[[2.564,-8.901,-1.981],[0.707106781,0,0,0.707106781],[0,0,0,0],[9E+09,9E+09,9E+09,9E+09,9E+09,9E+09]];
    CONST robtarget Target_Tap25_1050:=[[-25.909,-9.225,-2.248],[0.707106781,0,0,0.707106781],[0,0,0,0],[9E+09,9E+09,9E+09,9E+09,9E+09,9E+09]];
    CONST robtarget Target_Tap25_1060:=[[-25.909,-9.225,-20],[0.707106781,0,0,0.707106781],[0,0,0,0],[9E+09,9E+09,9E+09,9E+09,9E+09,9E+09]];
    CONST robtarget Target_Tap25_1070:=[[-31.985,-9.202,-20],[0.707106781,0,0,0.707106781],[0,0,0,0],[9E+09,9E+09,9E+09,9E+09,9E+09,9E+09]];
    CONST robtarget Target_Tap25_1080:=[[-31.981,-9.201,-2.285],[0.707106781,0,0,0.707106781],[0,0,0,0],[9E+09,9E+09,9E+09,9E+09,9E+09,9E+09]];
    CONST robtarget Target_Tap25_1090:=[[-40.518,-13.547,-2.372],[0.707106781,0,0,0.707106781],[0,0,0,0],[9E+09,9E+09,9E+09,9E+09,9E+09,9E+09]];
    CONST robtarget Target_Tap25_1100:=[[-47.252,-23.918,-2.433],[0.707106781,0,0,0.707106781],[0,0,0,0],[9E+09,9E+09,9E+09,9E+09,9E+09,9E+09]];
    CONST robtarget Target_Tap25_1110:=[[-47.252,-23.918,-20],[0.707106781,0,0,0.707106781],[0,0,0,0],[9E+09,9E+09,9E+09,9E+09,9E+09,9E+09]];
    CONST robtarget Target_Tap25_1120:=[[-46.96,-30.596,-20],[0.707106781,0,0,0.707106781],[0,0,0,0],[9E+09,9E+09,9E+09,9E+09,9E+09,9E+09]];
    CONST robtarget Target_Tap25_1130:=[[-46.96,-30.596,-2.43],[0.707106781,0,0,0.707106781],[0,0,0,0],[9E+09,9E+09,9E+09,9E+09,9E+09,9E+09]];
    CONST robtarget Target_Tap25_1140:=[[-41.363,-41.784,-2.38],[0.707106781,0,0,0.707106781],[0,0,0,0],[9E+09,9E+09,9E+09,9E+09,9E+09,9E+09]];
    CONST robtarget Target_Tap25_1150:=[[-31.622,-46.923,-2.282],[0.707106781,0,0,0.707106781],[0,0,0,0],[9E+09,9E+09,9E+09,9E+09,9E+09,9E+09]];
    CONST robtarget Target_Tap25_1160:=[[-31.622,-46.923,-20],[0.707106781,0,0,0.707106781],[0,0,0,0],[9E+09,9E+09,9E+09,9E+09,9E+09,9E+09]];
    CONST robtarget Target_Tap25_1170:=[[-26.538,-46.844,-20],[0.707106781,0,0,0.707106781],[0,0,0,0],[9E+09,9E+09,9E+09,9E+09,9E+09,9E+09]];
    CONST robtarget Target_Tap25_1180:=[[-26.538,-46.844,-2.254],[0.707106781,0,0,0.707106781],[0,0,0,0],[9E+09,9E+09,9E+09,9E+09,9E+09,9E+09]];
    CONST robtarget Target_Tap25_1190:=[[-16.389,-41.365,-2.153],[0.707106781,0,0,0.707106781],[0,0,0,0],[9E+09,9E+09,9E+09,9E+09,9E+09,9E+09]];
    CONST robtarget Target_Tap25_1200:=[[-11.855,-31.458,-2.112],[0.707106781,0,0,0.707106781],[0,0,0,0],[9E+09,9E+09,9E+09,9E+09,9E+09,9E+09]];
    CONST robtarget Target_Tap25_1210:=[[-11.759,-30.127,-20],[0.707106781,0,0,0.707106781],[0,0,0,0],[9E+09,9E+09,9E+09,9E+09,9E+09,9E+09]];
    CONST robtarget Target_Tap25_1220:=[[-29.396,-19.429,-20],[0.707106781,0,0,0.707106781],[0,0,0,0],[9E+09,9E+09,9E+09,9E+09,9E+09,9E+09]];
    CONST robtarget Target_Tap25_1230:=[[-29.396,-19.429,-2.271],[0.707106781,0,0,0.707106781],[0,0,0,0],[9E+09,9E+09,9E+09,9E+09,9E+09,9E+09]];
    CONST robtarget Target_Tap25_1240:=[[-26.364,-17.275,-2.243],[0.707106781,0,0,0.707106781],[0,0,0,0],[9E+09,9E+09,9E+09,9E+09,9E+09,9E+09]];
    CONST robtarget Target_Tap25_1250:=[[-23.419,-19.344,-2.217],[0.707106781,0,0,0.707106781],[0,0,0,0],[9E+09,9E+09,9E+09,9E+09,9E+09,9E+09]];
    CONST robtarget Target_Tap25_1260:=[[-24.634,-21.365,-2.228],[0.707106781,0,0,0.707106781],[0,0,0,0],[9E+09,9E+09,9E+09,9E+09,9E+09,9E+09]];
    CONST robtarget Target_Tap25_1270:=[[-29.583,-22.632,-2.273],[0.707106781,0,0,0.707106781],[0,0,0,0],[9E+09,9E+09,9E+09,9E+09,9E+09,9E+09]];
    CONST robtarget Target_Tap25_1280:=[[-26.708,-25.04,-2.247],[0.707106781,0,0,0.707106781],[0,0,0,0],[9E+09,9E+09,9E+09,9E+09,9E+09,9E+09]];
    CONST robtarget Target_Tap25_1290:=[[-23.233,-22.751,-2.215],[0.707106781,0,0,0.707106781],[0,0,0,0],[9E+09,9E+09,9E+09,9E+09,9E+09,9E+09]];
    CONST robtarget Target_Tap25_1300:=[[-23.233,-22.751,-20],[0.707106781,0,0,0.707106781],[0,0,0,0],[9E+09,9E+09,9E+09,9E+09,9E+09,9E+09]];
    CONST robtarget Target_Tap25_1310:=[[-18.61,-17.209,-20],[0.707106781,0,0,0.707106781],[0,0,0,0],[9E+09,9E+09,9E+09,9E+09,9E+09,9E+09]];
    CONST robtarget Target_Tap25_1320:=[[-18.61,-17.209,-2.173],[0.707106781,0,0,0.707106781],[0,0,0,0],[9E+09,9E+09,9E+09,9E+09,9E+09,9E+09]];
    CONST robtarget Target_Tap25_1330:=[[-22.347,-20.847,-2.207],[0.707106781,0,0,0.707106781],[0,0,0,0],[9E+09,9E+09,9E+09,9E+09,9E+09,9E+09]];
    CONST robtarget Target_Tap25_1340:=[[-18.674,-24.959,-2.174],[0.707106781,0,0,0.707106781],[0,0,0,0],[9E+09,9E+09,9E+09,9E+09,9E+09,9E+09]];
    CONST robtarget Target_Tap25_1350:=[[-14.796,-20.986,-2.138],[0.707106781,0,0,0.707106781],[0,0,0,0],[9E+09,9E+09,9E+09,9E+09,9E+09,9E+09]];
    CONST robtarget Target_Tap25_1360:=[[-18.654,-17.21,-2.173],[0.707106781,0,0,0.707106781],[0,0,0,0],[9E+09,9E+09,9E+09,9E+09,9E+09,9E+09]];
    CONST robtarget Target_Tap25_1370:=[[-18.654,-17.21,-20],[0.707106781,0,0,0.707106781],[0,0,0,0],[9E+09,9E+09,9E+09,9E+09,9E+09,9E+09]];
    CONST robtarget Target_Tap25_1380:=[[-13.597,-24.791,-20.128],[0.707106781,0,0,0.707106781],[0,0,0,0],[9E+09,9E+09,9E+09,9E+09,9E+09,9E+09]];
    CONST robtarget Target_Tap25_1390:=[[-13.597,-24.791,-2.128],[0.707106781,0,0,0.707106781],[0,0,0,0],[9E+09,9E+09,9E+09,9E+09,9E+09,9E+09]];
    CONST robtarget Target_Tap25_1400:=[[-13.578,-19.579,-2.127],[0.707106781,0,0,0.707106781],[0,0,0,0],[9E+09,9E+09,9E+09,9E+09,9E+09,9E+09]];
    CONST robtarget Target_Tap25_1410:=[[-11.844,-17.311,-2.112],[0.707106781,0,0,0.707106781],[0,0,0,0],[9E+09,9E+09,9E+09,9E+09,9E+09,9E+09]];
    CONST robtarget Target_Tap25_1420:=[[-8.417,-17.264,-2.081],[0.707106781,0,0,0.707106781],[0,0,0,0],[9E+09,9E+09,9E+09,9E+09,9E+09,9E+09]];
    CONST robtarget Target_Tap25_1430:=[[-7.647,-17.117,-2.074],[0.707106781,0,0,0.707106781],[0,0,0,0],[9E+09,9E+09,9E+09,9E+09,9E+09,9E+09]];
    CONST robtarget Target_Tap25_1440:=[[-7.427,-24.687,-2.072],[0.707106781,0,0,0.707106781],[0,0,0,0],[9E+09,9E+09,9E+09,9E+09,9E+09,9E+09]];
    CONST robtarget Target_Tap25_1450:=[[-7.446,-24.686,-20],[0.707106781,0,0,0.707106781],[0,0,0,0],[9E+09,9E+09,9E+09,9E+09,9E+09,9E+09]];
    CONST robtarget Target_Tap25_1460:=[[-7.635,-15.715,-20],[0.707106781,0,0,0.707106781],[0,0,0,0],[9E+09,9E+09,9E+09,9E+09,9E+09,9E+09]];
    CONST robtarget Target_Tap25_1470:=[[-7.635,-15.715,-0.073],[0.707106781,0,0,0.707106781],[0,0,0,0],[9E+09,9E+09,9E+09,9E+09,9E+09,9E+09]];
    CONST robtarget Target_Tap25_1480:=[[-9.976,-14.474,-0.095],[0.707106781,0,0,0.707106781],[0,0,0,0],[9E+09,9E+09,9E+09,9E+09,9E+09,9E+09]];
    CONST robtarget Target_Tap25_1490:=[[-11.372,-14.86,-0.107],[0.707106781,0,0,0.707106781],[0,0,0,0],[9E+09,9E+09,9E+09,9E+09,9E+09,9E+09]];
    CONST robtarget Target_Tap25_1500:=[[-12.954,-14.717,-0.122],[0.707106781,0,0,0.707106781],[0,0,0,0],[9E+09,9E+09,9E+09,9E+09,9E+09,9E+09]];
    CONST robtarget Target_Tap25_1510:=[[-12.954,-14.717,-20],[0.707106781,0,0,0.707106781],[0,0,0,0],[9E+09,9E+09,9E+09,9E+09,9E+09,9E+09]];
    CONST robtarget Target_Tap25_1520:=[[-3.81,-17.072,-20],[0.707106781,0,0,0.707106781],[0,0,0,0],[9E+09,9E+09,9E+09,9E+09,9E+09,9E+09]];
    CONST robtarget Target_Tap25_1530:=[[-3.81,-17.072,-2.039],[0.707106781,0,0,0.707106781],[0,0,0,0],[9E+09,9E+09,9E+09,9E+09,9E+09,9E+09]];
    CONST robtarget Target_Tap25_1540:=[[-3.921,-24.684,-2.04],[0.707106781,0,0,0.707106781],[0,0,0,0],[9E+09,9E+09,9E+09,9E+09,9E+09,9E+09]];
    CONST robtarget Target_Tap25_1550:=[[-2.602,-24.45,-2.028],[0.707106781,0,0,0.707106781],[0,0,0,0],[9E+09,9E+09,9E+09,9E+09,9E+09,9E+09]];
    CONST robtarget Target_Tap25_1560:=[[0.653,-24.611,-1.998],[0.707106781,0,0,0.707106781],[0,0,0,0],[9E+09,9E+09,9E+09,9E+09,9E+09,9E+09]];
    CONST robtarget Target_Tap25_1570:=[[2.916,-20.649,-1.978],[0.707106781,0,0,0.707106781],[0,0,0,0],[9E+09,9E+09,9E+09,9E+09,9E+09,9E+09]];
    CONST robtarget Target_Tap25_1580:=[[-0.061,-17.003,-2.005],[0.707106781,0,0,0.707106781],[0,0,0,0],[9E+09,9E+09,9E+09,9E+09,9E+09,9E+09]];
    CONST robtarget Target_Tap25_1590:=[[-2.661,-17.862,-2.028],[0.707106781,0,0,0.707106781],[0,0,0,0],[9E+09,9E+09,9E+09,9E+09,9E+09,9E+09]];
    CONST robtarget Target_Tap25_1600:=[[-2.661,-17.862,-20],[0.707106781,0,0,0.707106781],[0,0,0,0],[9E+09,9E+09,9E+09,9E+09,9E+09,9E+09]];
    CONST robtarget Target_Tap25_1610:=[[9.77,-34.658,-20],[0.707106781,0,0,0.707106781],[0,0,0,0],[9E+09,9E+09,9E+09,9E+09,9E+09,9E+09]];
    CONST robtarget Target_Tap25_1620:=[[9.728,-34.659,-1.934],[0.707106781,0,0,0.707106781],[0,0,0,0],[9E+09,9E+09,9E+09,9E+09,9E+09,9E+09]];
    CONST robtarget Target_Tap25_1630:=[[45.567,-34.033,-1.591],[0.707106781,0,0,0.707106781],[0,0,0,0],[9E+09,9E+09,9E+09,9E+09,9E+09,9E+09]];
    CONST robtarget Target_Tap25_1640:=[[34.516,-22.583,-1.7],[0.707106781,0,0,0.707106781],[0,0,0,0],[9E+09,9E+09,9E+09,9E+09,9E+09,9E+09]];
    CONST robtarget Target_Tap25_1650:=[[34.516,-22.583,-20],[0.707106781,0,0,0.707106781],[0,0,0,0],[9E+09,9E+09,9E+09,9E+09,9E+09,9E+09]];
    CONST robtarget Target_Tap25_1660:=[[30.036,-18.566,-20],[0.707106781,0,0,0.707106781],[0,0,0,0],[9E+09,9E+09,9E+09,9E+09,9E+09,9E+09]];
    CONST robtarget Target_Tap25_1670:=[[30.036,-18.566,-1.722],[0.707106781,0,0,0.707106781],[0,0,0,0],[9E+09,9E+09,9E+09,9E+09,9E+09,9E+09]];
    CONST robtarget Target_Tap25_1680:=[[9.182,6.895,-1.921],[0.707106781,0,0,0.707106781],[0,0,0,0],[9E+09,9E+09,9E+09,9E+09,9E+09,9E+09]];
    CONST robtarget Target_Tap25_1690:=[[20.558,40.249,-1.818],[0.707106781,0,0,0.707106781],[0,0,0,0],[9E+09,9E+09,9E+09,9E+09,9E+09,9E+09]];
    CONST robtarget Target_Tap25_1700:=[[40.908,46.872,-1.633],[0.707106781,0,0,0.707106781],[0,0,0,0],[9E+09,9E+09,9E+09,9E+09,9E+09,9E+09]];
    CONST robtarget Target_Tap25_1710:=[[64.938,35.959,-1.415],[0.707106781,0,0,0.707106781],[0,0,0,0],[9E+09,9E+09,9E+09,9E+09,9E+09,9E+09]];
    CONST robtarget Target_Tap25_1720:=[[72.742,14.835,-1.344],[0.707106781,0,0,0.707106781],[0,0,0,0],[9E+09,9E+09,9E+09,9E+09,9E+09,9E+09]];
    CONST robtarget Target_Tap25_1730:=[[72.773,14.835,-20],[0.707106781,0,0,0.707106781],[0,0,0,0],[9E+09,9E+09,9E+09,9E+09,9E+09,9E+09]];
    CONST robtarget Target_Tap25_1740:=[[62.787,14.87,-20],[0.707106781,0,0,0.707106781],[0,0,0,0],[9E+09,9E+09,9E+09,9E+09,9E+09,9E+09]];
    CONST robtarget Target_Tap25_1750:=[[62.787,14.87,-1.434],[0.707106781,0,0,0.707106781],[0,0,0,0],[9E+09,9E+09,9E+09,9E+09,9E+09,9E+09]];
    CONST robtarget Target_Tap25_1760:=[[56.474,30.558,-1.492],[0.707106781,0,0,0.707106781],[0,0,0,0],[9E+09,9E+09,9E+09,9E+09,9E+09,9E+09]];
    CONST robtarget Target_Tap25_1770:=[[42.723,36.93,-1.625],[0.707106781,0,0,0.707106781],[0,0,0,0],[9E+09,9E+09,9E+09,9E+09,9E+09,9E+09]];
    CONST robtarget Target_Tap25_1780:=[[42.723,36.93,-20],[0.707106781,0,0,0.707106781],[0,0,0,0],[9E+09,9E+09,9E+09,9E+09,9E+09,9E+09]];
    CONST robtarget Target_Tap25_1790:=[[38.707,36.257,-20],[0.707106781,0,0,0.707106781],[0,0,0,0],[9E+09,9E+09,9E+09,9E+09,9E+09,9E+09]];
    CONST robtarget Target_Tap25_1800:=[[37.707,36.257,-1.653],[0.707106781,0,0,0.707106781],[0,0,0,0],[9E+09,9E+09,9E+09,9E+09,9E+09,9E+09]];
    CONST robtarget Target_Tap25_1810:=[[23.045,30.043,-1.786],[0.707106781,0,0,0.707106781],[0,0,0,0],[9E+09,9E+09,9E+09,9E+09,9E+09,9E+09]];
    CONST robtarget Target_Tap25_1820:=[[18.351,16.476,-1.838],[0.707106781,0,0,0.707106781],[0,0,0,0],[9E+09,9E+09,9E+09,9E+09,9E+09,9E+09]];
    CONST robtarget Target_Tap25_1830:=[[18.351,16.476,-20],[0.707106781,0,0,0.707106781],[0,0,0,0],[9E+09,9E+09,9E+09,9E+09,9E+09,9E+09]];
    CONST robtarget Target_Tap25_1840:=[[18.267,10.708,-20],[0.707106781,0,0,0.707106781],[0,0,0,0],[9E+09,9E+09,9E+09,9E+09,9E+09,9E+09]];
    CONST robtarget Target_Tap25_1850:=[[18.267,10.708,-1.838],[0.707106781,0,0,0.707106781],[0,0,0,0],[9E+09,9E+09,9E+09,9E+09,9E+09,9E+09]];
    CONST robtarget Target_Tap25_1860:=[[21.963,2.727,-1.805],[0.707106781,0,0,0.707106781],[0,0,0,0],[9E+09,9E+09,9E+09,9E+09,9E+09,9E+09]];
    CONST robtarget Target_Tap25_1870:=[[36.377,-11.129,-1.665],[0.707106781,0,0,0.707106781],[0,0,0,0],[9E+09,9E+09,9E+09,9E+09,9E+09,9E+09]];
    CONST robtarget Target_Tap25_1880:=[[37.377,-12.129,-20],[0.707106781,0,0,0.707106781],[0,0,0,0],[9E+09,9E+09,9E+09,9E+09,9E+09,9E+09]];
    CONST robtarget Target_Tap25_1890:=[[40.514,-14.767,-20],[0.707106781,0,0,0.707106781],[0,0,0,0],[9E+09,9E+09,9E+09,9E+09,9E+09,9E+09]];
    CONST robtarget Target_Tap25_1900:=[[39.514,-13.767,-1.645],[0.707106781,0,0,0.707106781],[0,0,0,0],[9E+09,9E+09,9E+09,9E+09,9E+09,9E+09]];
    CONST robtarget Target_Tap25_1910:=[[50.447,-24.426,-1.546],[0.707106781,0,0,0.707106781],[0,0,0,0],[9E+09,9E+09,9E+09,9E+09,9E+09,9E+09]];
    CONST robtarget Target_Tap25_1920:=[[57.787,-33.113,-1.48],[0.707106781,0,0,0.707106781],[0,0,0,0],[9E+09,9E+09,9E+09,9E+09,9E+09,9E+09]];
    CONST robtarget Target_Tap25_1930:=[[63.784,-43.504,-1.425],[0.707106781,0,0,0.707106781],[0,0,0,0],[9E+09,9E+09,9E+09,9E+09,9E+09,9E+09]];
    CONST robtarget Target_Tap25_1940:=[[9.236,-44.416,-1.938],[0.707106781,0,0,0.707106781],[0,0,0,0],[9E+09,9E+09,9E+09,9E+09,9E+09,9E+09]];
    CONST robtarget Target_Tap25_1950:=[[9.236,-44.416,-20],[0.707106781,0,0,0.707106781],[0,0,0,0],[9E+09,9E+09,9E+09,9E+09,9E+09,9E+09]];
    CONST robtarget Target_Tap25_1960:=[[11.217,-62.22,-20],[0.707106781,0,0,0.707106781],[0,0,0,0],[9E+09,9E+09,9E+09,9E+09,9E+09,9E+09]];
    CONST robtarget Target_Tap25_1970:=[[11.217,-62.22,-1.902],[0.707106781,0,0,0.707106781],[0,0,0,0],[9E+09,9E+09,9E+09,9E+09,9E+09,9E+09]];
    CONST robtarget Target_Tap25_1980:=[[11.235,-68.995,-1.902],[0.707106781,0,0,0.707106781],[0,0,0,0],[9E+09,9E+09,9E+09,9E+09,9E+09,9E+09]];
    CONST robtarget Target_Tap25_1990:=[[12.22,-68.558,-1.893],[0.707106781,0,0,0.707106781],[0,0,0,0],[9E+09,9E+09,9E+09,9E+09,9E+09,9E+09]];
    CONST robtarget Target_Tap25_2000:=[[15.581,-68.844,-1.863],[0.707106781,0,0,0.707106781],[0,0,0,0],[9E+09,9E+09,9E+09,9E+09,9E+09,9E+09]];
    CONST robtarget Target_Tap25_2010:=[[17.244,-65.679,-1.848],[0.707106781,0,0,0.707106781],[0,0,0,0],[9E+09,9E+09,9E+09,9E+09,9E+09,9E+09]];
    CONST robtarget Target_Tap25_2020:=[[14.831,-62.1,-1.87],[0.707106781,0,0,0.707106781],[0,0,0,0],[9E+09,9E+09,9E+09,9E+09,9E+09,9E+09]];
    CONST robtarget Target_Tap25_2030:=[[12.402,-62.672,-1.892],[0.707106781,0,0,0.707106781],[0,0,0,0],[9E+09,9E+09,9E+09,9E+09,9E+09,9E+09]];
    CONST robtarget Target_Tap25_2040:=[[12.402,-62.672,-20],[0.707106781,0,0,0.707106781],[0,0,0,0],[9E+09,9E+09,9E+09,9E+09,9E+09,9E+09]];
    CONST robtarget Target_Tap25_2050:=[[19.743,-68.941,-20],[0.707106781,0,0,0.707106781],[0,0,0,0],[9E+09,9E+09,9E+09,9E+09,9E+09,9E+09]];
    CONST robtarget Target_Tap25_2060:=[[19.77,-68.941,-1.825],[0.707106781,0,0,0.707106781],[0,0,0,0],[9E+09,9E+09,9E+09,9E+09,9E+09,9E+09]];
    CONST robtarget Target_Tap25_2070:=[[19.573,-62.094,-1.826],[0.707106781,0,0,0.707106781],[0,0,0,0],[9E+09,9E+09,9E+09,9E+09,9E+09,9E+09]];
    CONST robtarget Target_Tap25_2080:=[[19.628,-62.094,-20],[0.707106781,0,0,0.707106781],[0,0,0,0],[9E+09,9E+09,9E+09,9E+09,9E+09,9E+09]];
    CONST robtarget Target_Tap25_2090:=[[20.869,-60.282,-20],[0.707106781,0,0,0.707106781],[0,0,0,0],[9E+09,9E+09,9E+09,9E+09,9E+09,9E+09]];
    CONST robtarget Target_Tap25_2100:=[[20.864,-59.882,-1.815],[0.707106781,0,0,0.707106781],[0,0,0,0],[9E+09,9E+09,9E+09,9E+09,9E+09,9E+09]];
    CONST robtarget Target_Tap25_2110:=[[17.984,-59.006,-1.841],[0.707106781,0,0,0.707106781],[0,0,0,0],[9E+09,9E+09,9E+09,9E+09,9E+09,9E+09]];
    CONST robtarget Target_Tap25_2120:=[[17.984,-59.006,-20],[0.707106781,0,0,0.707106781],[0,0,0,0],[9E+09,9E+09,9E+09,9E+09,9E+09,9E+09]];
    CONST robtarget Target_Tap25_2130:=[[21.806,-63.077,-20],[0.707106781,0,0,0.707106781],[0,0,0,0],[9E+09,9E+09,9E+09,9E+09,9E+09,9E+09]];
    CONST robtarget Target_Tap25_2140:=[[21.806,-63.077,0.194],[0.707106781,0,0,0.707106781],[0,0,0,0],[9E+09,9E+09,9E+09,9E+09,9E+09,9E+09]];
    CONST robtarget Target_Tap25_2150:=[[23.747,-62.749,-1.789],[0.707106781,0,0,0.707106781],[0,0,0,0],[9E+09,9E+09,9E+09,9E+09,9E+09,9E+09]];
    CONST robtarget Target_Tap25_2160:=[[24.9,-62.036,-1.778],[0.707106781,0,0,0.707106781],[0,0,0,0],[9E+09,9E+09,9E+09,9E+09,9E+09,9E+09]];
    CONST robtarget Target_Tap25_2170:=[[25.062,-68.782,-1.777],[0.707106781,0,0,0.707106781],[0,0,0,0],[9E+09,9E+09,9E+09,9E+09,9E+09,9E+09]];
    CONST robtarget Target_Tap25_2180:=[[25.062,-68.782,-20],[0.707106781,0,0,0.707106781],[0,0,0,0],[9E+09,9E+09,9E+09,9E+09,9E+09,9E+09]];
    CONST robtarget Target_Tap25_2190:=[[27.285,-66.763,-20],[0.707106781,0,0,0.707106781],[0,0,0,0],[9E+09,9E+09,9E+09,9E+09,9E+09,9E+09]];
    CONST robtarget Target_Tap25_2200:=[[27.285,-66.763,-1.756],[0.707106781,0,0,0.707106781],[0,0,0,0],[9E+09,9E+09,9E+09,9E+09,9E+09,9E+09]];
    CONST robtarget Target_Tap25_2210:=[[30.688,-68.964,-1.726],[0.707106781,0,0,0.707106781],[0,0,0,0],[9E+09,9E+09,9E+09,9E+09,9E+09,9E+09]];
    CONST robtarget Target_Tap25_2220:=[[33.804,-65.581,-1.697],[0.707106781,0,0,0.707106781],[0,0,0,0],[9E+09,9E+09,9E+09,9E+09,9E+09,9E+09]];
    CONST robtarget Target_Tap25_2230:=[[30.598,-61.876,-1.726],[0.707106781,0,0,0.707106781],[0,0,0,0],[9E+09,9E+09,9E+09,9E+09,9E+09,9E+09]];
    CONST robtarget Target_Tap25_2240:=[[27.073,-65.839,-1.758],[0.707106781,0,0,0.707106781],[0,0,0,0],[9E+09,9E+09,9E+09,9E+09,9E+09,9E+09]];
    CONST robtarget Target_Tap25_2250:=[[31.649,-65.959,-1.717],[0.707106781,0,0,0.707106781],[0,0,0,0],[9E+09,9E+09,9E+09,9E+09,9E+09,9E+09]];
    CONST robtarget Target_Tap25_2260:=[[31.649,-65.959,-20],[0.707106781,0,0,0.707106781],[0,0,0,0],[9E+09,9E+09,9E+09,9E+09,9E+09,9E+09]];
    CONST robtarget Target_Tap25_2270:=[[36.079,-68.725,-20],[0.707106781,0,0,0.707106781],[0,0,0,0],[9E+09,9E+09,9E+09,9E+09,9E+09,9E+09]];
    CONST robtarget Target_Tap25_2280:=[[36.079,-68.725,-1.677],[0.707106781,0,0,0.707106781],[0,0,0,0],[9E+09,9E+09,9E+09,9E+09,9E+09,9E+09]];
    CONST robtarget Target_Tap25_2290:=[[35.934,-61.955,-1.678],[0.707106781,0,0,0.707106781],[0,0,0,0],[9E+09,9E+09,9E+09,9E+09,9E+09,9E+09]];
    CONST robtarget Target_Tap25_2300:=[[35.934,-61.955,-20],[0.707106781,0,0,0.707106781],[0,0,0,0],[9E+09,9E+09,9E+09,9E+09,9E+09,9E+09]];
    CONST robtarget Target_Tap25_2310:=[[39.604,-68.678,-20],[0.707106781,0,0,0.707106781],[0,0,0,0],[9E+09,9E+09,9E+09,9E+09,9E+09,9E+09]];
    CONST robtarget Target_Tap25_2320:=[[39.604,-68.678,-1.645],[0.707106781,0,0,0.707106781],[0,0,0,0],[9E+09,9E+09,9E+09,9E+09,9E+09,9E+09]];
    CONST robtarget Target_Tap25_2330:=[[39.562,-62.217,-1.645],[0.707106781,0,0,0.707106781],[0,0,0,0],[9E+09,9E+09,9E+09,9E+09,9E+09,9E+09]];
    CONST robtarget Target_Tap25_2340:=[[43.112,-62.258,-1.613],[0.707106781,0,0,0.707106781],[0,0,0,0],[9E+09,9E+09,9E+09,9E+09,9E+09,9E+09]];
    CONST robtarget Target_Tap25_2350:=[[44.045,-61.827,-1.604],[0.707106781,0,0,0.707106781],[0,0,0,0],[9E+09,9E+09,9E+09,9E+09,9E+09,9E+09]];
    CONST robtarget Target_Tap25_2360:=[[44.225,-68.672,-1.603],[0.707106781,0,0,0.707106781],[0,0,0,0],[9E+09,9E+09,9E+09,9E+09,9E+09,9E+09]];
    CONST robtarget Target_Tap25_2370:=[[44.225,-68.672,-20],[0.707106781,0,0,0.707106781],[0,0,0,0],[9E+09,9E+09,9E+09,9E+09,9E+09,9E+09]];
    CONST robtarget Target_Tap25_2380:=[[46.488,-66.774,-20],[0.707106781,0,0,0.707106781],[0,0,0,0],[9E+09,9E+09,9E+09,9E+09,9E+09,9E+09]];
    CONST robtarget Target_Tap25_2390:=[[46.488,-66.774,-1.582],[0.707106781,0,0,0.707106781],[0,0,0,0],[9E+09,9E+09,9E+09,9E+09,9E+09,9E+09]];
    CONST robtarget Target_Tap25_2400:=[[49.146,-68.737,-1.558],[0.707106781,0,0,0.707106781],[0,0,0,0],[9E+09,9E+09,9E+09,9E+09,9E+09,9E+09]];
    CONST robtarget Target_Tap25_2410:=[[52.369,-67.36,-1.529],[0.707106781,0,0,0.707106781],[0,0,0,0],[9E+09,9E+09,9E+09,9E+09,9E+09,9E+09]];
    CONST robtarget Target_Tap25_2420:=[[51.363,-62.022,-1.538],[0.707106781,0,0,0.707106781],[0,0,0,0],[9E+09,9E+09,9E+09,9E+09,9E+09,9E+09]];
    CONST robtarget Target_Tap25_2430:=[[46.186,-65.629,-1.585],[0.707106781,0,0,0.707106781],[0,0,0,0],[9E+09,9E+09,9E+09,9E+09,9E+09,9E+09]];
    CONST robtarget Target_Tap25_2440:=[[50.972,-65.902,-1.542],[0.707106781,0,0,0.707106781],[0,0,0,0],[9E+09,9E+09,9E+09,9E+09,9E+09,9E+09]];
    CONST robtarget Target_Tap25_2450:=[[50.972,-65.902,-20],[0.707106781,0,0,0.707106781],[0,0,0,0],[9E+09,9E+09,9E+09,9E+09,9E+09,9E+09]];
    CONST robtarget Target_Tap25_2460:=[[60.95,-69.621,-20],[0.707106781,0,0,0.707106781],[0,0,0,0],[9E+09,9E+09,9E+09,9E+09,9E+09,9E+09]];
    CONST robtarget Target_Tap25_2470:=[[60.95,-69.621,-1.451],[0.707106781,0,0,0.707106781],[0,0,0,0],[9E+09,9E+09,9E+09,9E+09,9E+09,9E+09]];
    CONST robtarget Target_Tap25_2480:=[[57.957,-71.923,-1.478],[0.707106781,0,0,0.707106781],[0,0,0,0],[9E+09,9E+09,9E+09,9E+09,9E+09,9E+09]];
    CONST robtarget Target_Tap25_2490:=[[54.509,-69.871,-1.509],[0.707106781,0,0,0.707106781],[0,0,0,0],[9E+09,9E+09,9E+09,9E+09,9E+09,9E+09]];
    CONST robtarget Target_Tap25_2500:=[[54.222,-61.87,-1.512],[0.707106781,0,0,0.707106781],[0,0,0,0],[9E+09,9E+09,9E+09,9E+09,9E+09,9E+09]];
    CONST robtarget Target_Tap25_2510:=[[56.097,-61.975,-1.495],[0.707106781,0,0,0.707106781],[0,0,0,0],[9E+09,9E+09,9E+09,9E+09,9E+09,9E+09]];
    CONST robtarget Target_Tap25_2520:=[[59.946,-62.085,-1.46],[0.707106781,0,0,0.707106781],[0,0,0,0],[9E+09,9E+09,9E+09,9E+09,9E+09,9E+09]];
    CONST robtarget Target_Tap25_2530:=[[61.014,-66.567,-1.45],[0.707106781,0,0,0.707106781],[0,0,0,0],[9E+09,9E+09,9E+09,9E+09,9E+09,9E+09]];
    CONST robtarget Target_Tap25_2540:=[[56.657,-68.05,-1.49],[0.707106781,0,0,0.707106781],[0,0,0,0],[9E+09,9E+09,9E+09,9E+09,9E+09,9E+09]];
    CONST robtarget Target_Tap25_2550:=[[56.657,-68.05,-20],[0.707106781,0,0,0.707106781],[0,0,0,0],[9E+09,9E+09,9E+09,9E+09,9E+09,9E+09]];
    CONST robtarget Target_Tap25_2560:=[[63.194,-68.464,-19.431],[0.707106781,0,0,0.707106781],[0,0,0,0],[9E+09,9E+09,9E+09,9E+09,9E+09,9E+09]];
    CONST robtarget Target_Tap25_2570:=[[63.194,-68.464,-1.431],[0.707106781,0,0,0.707106781],[0,0,0,0],[9E+09,9E+09,9E+09,9E+09,9E+09,9E+09]];
    CONST robtarget Target_Tap25_2580:=[[63.388,-61.935,-1.429],[0.707106781,0,0,0.707106781],[0,0,0,0],[9E+09,9E+09,9E+09,9E+09,9E+09,9E+09]];
    CONST robtarget Target_Tap25_2590:=[[66.746,-62.021,-1.398],[0.707106781,0,0,0.707106781],[0,0,0,0],[9E+09,9E+09,9E+09,9E+09,9E+09,9E+09]];
    CONST robtarget Target_Tap25_2600:=[[67.896,-61.563,-1.388],[0.707106781,0,0,0.707106781],[0,0,0,0],[9E+09,9E+09,9E+09,9E+09,9E+09,9E+09]];
    CONST robtarget Target_Tap25_2610:=[[67.926,-68.412,-1.388],[0.707106781,0,0,0.707106781],[0,0,0,0],[9E+09,9E+09,9E+09,9E+09,9E+09,9E+09]];
    CONST robtarget Target_Tap25_2620:=[[67.926,-68.412,-20],[0.707106781,0,0,0.707106781],[0,0,0,0],[9E+09,9E+09,9E+09,9E+09,9E+09,9E+09]];
    CONST robtarget Target_Tap25_2630:=[[71.585,-68.371,-20],[0.707106781,0,0,0.707106781],[0,0,0,0],[9E+09,9E+09,9E+09,9E+09,9E+09,9E+09]];
    CONST robtarget Target_Tap25_2640:=[[71.585,-68.371,-1.354],[0.707106781,0,0,0.707106781],[0,0,0,0],[9E+09,9E+09,9E+09,9E+09,9E+09,9E+09]];
    CONST robtarget Target_Tap25_2650:=[[71.464,-59.512,-1.356],[0.707106781,0,0,0.707106781],[0,0,0,0],[9E+09,9E+09,9E+09,9E+09,9E+09,9E+09]];
    CONST robtarget Target_Tap25_2660:=[[71.464,-59.512,-20],[0.707106781,0,0,0.707106781],[0,0,0,0],[9E+09,9E+09,9E+09,9E+09,9E+09,9E+09]];
    CONST robtarget Target_Tap25_2670:=[[75.802,61.109,-20],[0.707106781,0,0,0.707106781],[0,0,0,0],[9E+09,9E+09,9E+09,9E+09,9E+09,9E+09]];
    CONST robtarget Target_Tap25_2680:=[[75.802,61.109,-1.316],[0.707106781,0,0,0.707106781],[0,0,0,0],[9E+09,9E+09,9E+09,9E+09,9E+09,9E+09]];
    CONST robtarget Target_Tap25_2690:=[[74.944,70.264,-1.324],[0.707106781,0,0,0.707106781],[0,0,0,0],[9E+09,9E+09,9E+09,9E+09,9E+09,9E+09]];
    CONST robtarget Target_Tap25_2700:=[[67.504,69.191,-1.391],[0.707106781,0,0,0.707106781],[0,0,0,0],[9E+09,9E+09,9E+09,9E+09,9E+09,9E+09]];
    CONST robtarget Target_Tap25_2710:=[[70.964,51.233,-1.36],[0.707106781,0,0,0.707106781],[0,0,0,0],[9E+09,9E+09,9E+09,9E+09,9E+09,9E+09]];
    CONST robtarget Target_Tap25_2720:=[[59.916,59.844,-1.46],[0.707106781,0,0,0.707106781],[0,0,0,0],[9E+09,9E+09,9E+09,9E+09,9E+09,9E+09]];
    CONST robtarget Target_Tap25_2730:=[[59.931,59.865,-20],[0.707106781,0,0,0.707106781],[0,0,0,0],[9E+09,9E+09,9E+09,9E+09,9E+09,9E+09]];
    CONST robtarget Target_Tap25_2740:=[[49.511,63.12,-20],[0.707106781,0,0,0.707106781],[0,0,0,0],[9E+09,9E+09,9E+09,9E+09,9E+09,9E+09]];
    CONST robtarget Target_Tap25_2750:=[[49.508,63.121,-1.555],[0.707106781,0,0,0.707106781],[0,0,0,0],[9E+09,9E+09,9E+09,9E+09,9E+09,9E+09]];
    CONST robtarget Target_Tap25_2760:=[[60.017,67.312,-1.459],[0.707106781,0,0,0.707106781],[0,0,0,0],[9E+09,9E+09,9E+09,9E+09,9E+09,9E+09]];
    CONST robtarget Target_Tap25_2770:=[[57.983,80.74,-1.478],[0.707106781,0,0,0.707106781],[0,0,0,0],[9E+09,9E+09,9E+09,9E+09,9E+09,9E+09]];
    CONST robtarget Target_Tap25_2780:=[[46.809,75.946,-1.579],[0.707106781,0,0,0.707106781],[0,0,0,0],[9E+09,9E+09,9E+09,9E+09,9E+09,9E+09]];
    CONST robtarget Target_Tap25_2790:=[[49.544,63.101,-1.554],[0.707106781,0,0,0.707106781],[0,0,0,0],[9E+09,9E+09,9E+09,9E+09,9E+09,9E+09]];
    CONST robtarget Target_Tap25_2800:=[[49.505,63.123,-20],[0.707106781,0,0,0.707106781],[0,0,0,0],[9E+09,9E+09,9E+09,9E+09,9E+09,9E+09]];
    CONST robtarget Target_Tap25_2810:=[[31.853,70.292,-20],[0.707106781,0,0,0.707106781],[0,0,0,0],[9E+09,9E+09,9E+09,9E+09,9E+09,9E+09]];
    CONST robtarget Target_Tap25_2820:=[[31.85,70.293,-1.715],[0.707106781,0,0,0.707106781],[0,0,0,0],[9E+09,9E+09,9E+09,9E+09,9E+09,9E+09]];
    CONST robtarget Target_Tap25_2830:=[[41.877,77.147,-1.624],[0.707106781,0,0,0.707106781],[0,0,0,0],[9E+09,9E+09,9E+09,9E+09,9E+09,9E+09]];
    CONST robtarget Target_Tap25_2840:=[[37.197,89.053,-1.667],[0.707106781,0,0,0.707106781],[0,0,0,0],[9E+09,9E+09,9E+09,9E+09,9E+09,9E+09]];
    CONST robtarget Target_Tap25_2850:=[[26.745,81.247,-1.761],[0.707106781,0,0,0.707106781],[0,0,0,0],[9E+09,9E+09,9E+09,9E+09,9E+09,9E+09]];
    CONST robtarget Target_Tap25_2860:=[[31.814,70.304,-1.715],[0.707106781,0,0,0.707106781],[0,0,0,0],[9E+09,9E+09,9E+09,9E+09,9E+09,9E+09]];
    CONST robtarget Target_Tap25_2870:=[[31.814,70.304,-20],[0.707106781,0,0,0.707106781],[0,0,0,0],[9E+09,9E+09,9E+09,9E+09,9E+09,9E+09]];
    CONST robtarget Target_Tap25_2880:=[[15.701,73.888,-20],[0.707106781,0,0,0.707106781],[0,0,0,0],[9E+09,9E+09,9E+09,9E+09,9E+09,9E+09]];
    CONST robtarget Target_Tap25_2890:=[[15.734,73.884,-1.861],[0.707106781,0,0,0.707106781],[0,0,0,0],[9E+09,9E+09,9E+09,9E+09,9E+09,9E+09]];
    CONST robtarget Target_Tap25_2900:=[[18.684,92.872,-1.835],[0.707106781,0,0,0.707106781],[0,0,0,0],[9E+09,9E+09,9E+09,9E+09,9E+09,9E+09]];
    CONST robtarget Target_Tap25_2910:=[[23.889,91.77,-1.787],[0.707106781,0,0,0.707106781],[0,0,0,0],[9E+09,9E+09,9E+09,9E+09,9E+09,9E+09]];
    CONST robtarget Target_Tap25_2920:=[[23.889,91.77,-20],[0.707106781,0,0,0.707106781],[0,0,0,0],[9E+09,9E+09,9E+09,9E+09,9E+09,9E+09]];
    CONST robtarget Target_Tap25_2930:=[[8.703,84.352,-20],[0.707106781,0,0,0.707106781],[0,0,0,0],[9E+09,9E+09,9E+09,9E+09,9E+09,9E+09]];
    CONST robtarget Target_Tap25_2940:=[[8.703,84.352,-1.925],[0.707106781,0,0,0.707106781],[0,0,0,0],[9E+09,9E+09,9E+09,9E+09,9E+09,9E+09]];
    CONST robtarget Target_Tap25_2950:=[[-3.378,83.892,-2.035],[0.707106781,0,0,0.707106781],[0,0,0,0],[9E+09,9E+09,9E+09,9E+09,9E+09,9E+09]];
    CONST robtarget Target_Tap25_2960:=[[-3.378,83.892,-20],[0.707106781,0,0,0.707106781],[0,0,0,0],[9E+09,9E+09,9E+09,9E+09,9E+09,9E+09]];
    CONST robtarget Target_Tap25_2970:=[[-12.295,87.107,-20],[0.707106781,0,0,0.707106781],[0,0,0,0],[9E+09,9E+09,9E+09,9E+09,9E+09,9E+09]];
    CONST robtarget Target_Tap25_2980:=[[-12.295,87.107,-2.116],[0.707106781,0,0,0.707106781],[0,0,0,0],[9E+09,9E+09,9E+09,9E+09,9E+09,9E+09]];
    CONST robtarget Target_Tap25_2990:=[[-17.721,93.248,-2.165],[0.707106781,0,0,0.707106781],[0,0,0,0],[9E+09,9E+09,9E+09,9E+09,9E+09,9E+09]];
    CONST robtarget Target_Tap25_3000:=[[-23.929,87.687,-2.221],[0.707106781,0,0,0.707106781],[0,0,0,0],[9E+09,9E+09,9E+09,9E+09,9E+09,9E+09]];
    CONST robtarget Target_Tap25_3010:=[[-8.74,77.04,-2.083],[0.707106781,0,0,0.707106781],[0,0,0,0],[9E+09,9E+09,9E+09,9E+09,9E+09,9E+09]];
    CONST robtarget Target_Tap25_3020:=[[-22.719,75.151,-2.21],[0.707106781,0,0,0.707106781],[0,0,0,0],[9E+09,9E+09,9E+09,9E+09,9E+09,9E+09]];
    CONST robtarget Target_Tap25_3030:=[[-22.707,75.082,-20],[0.707106781,0,0,0.707106781],[0,0,0,0],[9E+09,9E+09,9E+09,9E+09,9E+09,9E+09]];
    CONST robtarget Target_Tap25_3040:=[[-32.775,69.883,-20],[0.707106781,0,0,0.707106781],[0,0,0,0],[9E+09,9E+09,9E+09,9E+09,9E+09,9E+09]];
    CONST robtarget Target_Tap25_3050:=[[-32.74,69.893,-2.301],[0.707106781,0,0,0.707106781],[0,0,0,0],[9E+09,9E+09,9E+09,9E+09,9E+09,9E+09]];
    CONST robtarget Target_Tap25_3060:=[[-28.406,82.137,-2.262],[0.707106781,0,0,0.707106781],[0,0,0,0],[9E+09,9E+09,9E+09,9E+09,9E+09,9E+09]];
    CONST robtarget Target_Tap25_3070:=[[-38.484,88.525,-2.353],[0.707106781,0,0,0.707106781],[0,0,0,0],[9E+09,9E+09,9E+09,9E+09,9E+09,9E+09]];
    CONST robtarget Target_Tap25_3080:=[[-43.532,78.171,-2.399],[0.707106781,0,0,0.707106781],[0,0,0,0],[9E+09,9E+09,9E+09,9E+09,9E+09,9E+09]];
    CONST robtarget Target_Tap25_3090:=[[-32.74,69.893,-2.301],[0.707106781,0,0,0.707106781],[0,0,0,0],[9E+09,9E+09,9E+09,9E+09,9E+09,9E+09]];
    CONST robtarget Target_Tap25_3100:=[[-32.74,69.893,-20],[0.707106781,0,0,0.707106781],[0,0,0,0],[9E+09,9E+09,9E+09,9E+09,9E+09,9E+09]];
    CONST robtarget Target_Tap25_3110:=[[-51.172,76.399,-20],[0.707106781,0,0,0.707106781],[0,0,0,0],[9E+09,9E+09,9E+09,9E+09,9E+09,9E+09]];
    CONST robtarget Target_Tap25_3120:=[[-51.143,76.415,-2.468],[0.707106781,0,0,0.707106781],[0,0,0,0],[9E+09,9E+09,9E+09,9E+09,9E+09,9E+09]];
    CONST robtarget Target_Tap25_3130:=[[-59.237,79.994,-2.542],[0.707106781,0,0,0.707106781],[0,0,0,0],[9E+09,9E+09,9E+09,9E+09,9E+09,9E+09]];
    CONST robtarget Target_Tap25_3140:=[[-62.202,73.588,-2.569],[0.707106781,0,0,0.707106781],[0,0,0,0],[9E+09,9E+09,9E+09,9E+09,9E+09,9E+09]];
    CONST robtarget Target_Tap25_3150:=[[-44.322,68.42,-2.406],[0.707106781,0,0,0.707106781],[0,0,0,0],[9E+09,9E+09,9E+09,9E+09,9E+09,9E+09]];
    CONST robtarget Target_Tap25_3160:=[[-56.604,61.373,-2.518],[0.707106781,0,0,0.707106781],[0,0,0,0],[9E+09,9E+09,9E+09,9E+09,9E+09,9E+09]];
    CONST robtarget Target_Tap25_3170:=[[-56.604,61.373,-20],[0.707106781,0,0,0.707106781],[0,0,0,0],[9E+09,9E+09,9E+09,9E+09,9E+09,9E+09]];
    CONST robtarget Target_Tap25_3180:=[[-76.573,61.848,-20],[0.707106781,0,0,0.707106781],[0,0,0,0],[9E+09,9E+09,9E+09,9E+09,9E+09,9E+09]];
    CONST robtarget Target_Tap25_3190:=[[-76.573,61.848,-2.699],[0.707106781,0,0,0.707106781],[0,0,0,0],[9E+09,9E+09,9E+09,9E+09,9E+09,9E+09]];
    CONST robtarget Target_Tap25_3200:=[[-75.943,69.496,-2.693],[0.707106781,0,0,0.707106781],[0,0,0,0],[9E+09,9E+09,9E+09,9E+09,9E+09,9E+09]];
    CONST robtarget Target_Tap25_3210:=[[-66.167,67.964,-2.605],[0.707106781,0,0,0.707106781],[0,0,0,0],[9E+09,9E+09,9E+09,9E+09,9E+09,9E+09]];
    CONST robtarget Target_Tap25_3220:=[[-61.498,57.083,-2.562],[0.707106781,0,0,0.707106781],[0,0,0,0],[9E+09,9E+09,9E+09,9E+09,9E+09,9E+09]];
    CONST robtarget Target_Tap25_3230:=[[-65.646,52.346,-2.6],[0.707106781,0,0,0.707106781],[0,0,0,0],[9E+09,9E+09,9E+09,9E+09,9E+09,9E+09]];
    CONST robtarget Target_Tap25_3240:=[[-73.893,54.168,-2.675],[0.707106781,0,0,0.707106781],[0,0,0,0],[9E+09,9E+09,9E+09,9E+09,9E+09,9E+09]];
    CONST robtarget Target_Tap25_3250:=[[-73.022,62.517,-2.667],[0.707106781,0,0,0.707106781],[0,0,0,0],[9E+09,9E+09,9E+09,9E+09,9E+09,9E+09]];
    CONST robtarget Target_Tap25_3260:=[[-64.723,66.076,-2.628],[0.707106781,0,0,0.707106781],[0,0,0,0],[9E+09,9E+09,9E+09,9E+09,9E+09,9E+09]];
    CONST robtarget Target_Tap25_3270:=[[-68.896,64.06,-20],[0.707106781,0,0,0.707106781],[0,0,0,0],[9E+09,9E+09,9E+09,9E+09,9E+09,9E+09]];
    CONST robtarget p_contacto_25{279}:=[Target_Tap25_20, Target_Tap25_30, Target_Tap25_40, Target_Tap25_50, Target_Tap25_60, Target_Tap25_70,
                                      Target_Tap25_90, Target_Tap25_100, Target_Tap25_110, Target_Tap25_120, Target_Tap25_130, Target_Tap25_140,
                                      Target_Tap25_150, Target_Tap25_170, Target_Tap25_180, Target_Tap25_190, Target_Tap25_200, Target_Tap25_210,
                                      Target_Tap25_220, Target_Tap25_240, Target_Tap25_250, Target_Tap25_260, Target_Tap25_270, Target_Tap25_280,
                                      Target_Tap25_290, Target_Tap25_300, Target_Tap25_310, Target_Tap25_320, Target_Tap25_340, Target_Tap25_350,
                                      Target_Tap25_360, Target_Tap25_370, Target_Tap25_380, Target_Tap25_390, Target_Tap25_400, Target_Tap25_410,
                                      Target_Tap25_420, Target_Tap25_440, Target_Tap25_450, Target_Tap25_460, Target_Tap25_470, Target_Tap25_480,
                                      Target_Tap25_500, Target_Tap25_510, Target_Tap25_520, Target_Tap25_540, Target_Tap25_550, Target_Tap25_560,
                                      Target_Tap25_570, Target_Tap25_580, Target_Tap25_590, Target_Tap25_610, Target_Tap25_620, Target_Tap25_630,
                                      Target_Tap25_640, Target_Tap25_650, Target_Tap25_660, Target_Tap25_670, Target_Tap25_690, Target_Tap25_700,
                                      Target_Tap25_710, Target_Tap25_730, Target_Tap25_740, Target_Tap25_760, Target_Tap25_770, Target_Tap25_780,
                                      Target_Tap25_790, Target_Tap25_800, Target_Tap25_810, Target_Tap25_830, Target_Tap25_840, Target_Tap25_850,
                                      Target_Tap25_860, Target_Tap25_870, Target_Tap25_880, Target_Tap25_890, Target_Tap25_900, Target_Tap25_920,
                                      Target_Tap25_930, Target_Tap25_940, Target_Tap25_950, Target_Tap25_960, Target_Tap25_970, Target_Tap25_980,
                                      Target_Tap25_990, Target_Tap25_1000, Target_Tap25_1020, Target_Tap25_1030, Target_Tap25_1040, Target_Tap25_1050,
                                      Target_Tap25_1060, Target_Tap25_1080, Target_Tap25_1090, Target_Tap25_1100, Target_Tap25_1110, Target_Tap25_1130,
                                      Target_Tap25_1140, Target_Tap25_1150, Target_Tap25_1160, Target_Tap25_1180, Target_Tap25_1190, Target_Tap25_1200,
                                      Target_Tap25_1210, Target_Tap25_1230, Target_Tap25_1240, Target_Tap25_1250, Target_Tap25_1260, Target_Tap25_1270,
                                      Target_Tap25_1280, Target_Tap25_1290, Target_Tap25_1300, Target_Tap25_1320, Target_Tap25_1330, Target_Tap25_1340,
                                      Target_Tap25_1350, Target_Tap25_1360, Target_Tap25_1370, Target_Tap25_1390, Target_Tap25_1400, Target_Tap25_1410,
                                      Target_Tap25_1420, Target_Tap25_1430, Target_Tap25_1440, Target_Tap25_1450, Target_Tap25_1470, Target_Tap25_1480,
                                      Target_Tap25_1490, Target_Tap25_1500, Target_Tap25_1510, Target_Tap25_1530, Target_Tap25_1540, Target_Tap25_1550,
                                      Target_Tap25_1560, Target_Tap25_1570, Target_Tap25_1580, Target_Tap25_1590, Target_Tap25_1600, Target_Tap25_1620,
                                      Target_Tap25_1630, Target_Tap25_1640, Target_Tap25_1650, Target_Tap25_1670, Target_Tap25_1680, Target_Tap25_1690,
                                      Target_Tap25_1700, Target_Tap25_1710, Target_Tap25_1720, Target_Tap25_1730, Target_Tap25_1750, Target_Tap25_1760,
                                      Target_Tap25_1770, Target_Tap25_1780, Target_Tap25_1800, Target_Tap25_1810, Target_Tap25_1820, Target_Tap25_1830,
                                      Target_Tap25_1850, Target_Tap25_1860, Target_Tap25_1870, Target_Tap25_1880, Target_Tap25_1900, Target_Tap25_1910,
                                      Target_Tap25_1920, Target_Tap25_1930, Target_Tap25_1940, Target_Tap25_1950, Target_Tap25_1970, Target_Tap25_1980,
                                      Target_Tap25_1990, Target_Tap25_2000, Target_Tap25_2010, Target_Tap25_2020, Target_Tap25_2030, Target_Tap25_2040,
                                      Target_Tap25_2060, Target_Tap25_2070, Target_Tap25_2080, Target_Tap25_2100, Target_Tap25_2110, Target_Tap25_2120,
                                      Target_Tap25_2140, Target_Tap25_2150, Target_Tap25_2160, Target_Tap25_2170, Target_Tap25_2180, Target_Tap25_2200,
                                      Target_Tap25_2210, Target_Tap25_2220, Target_Tap25_2230, Target_Tap25_2240, Target_Tap25_2250, Target_Tap25_2260,
                                      Target_Tap25_2280, Target_Tap25_2290, Target_Tap25_2300, Target_Tap25_2320, Target_Tap25_2330, Target_Tap25_2340,
                                      Target_Tap25_2350, Target_Tap25_2360, Target_Tap25_2370, Target_Tap25_2390, Target_Tap25_2400, Target_Tap25_2410,
                                      Target_Tap25_2420, Target_Tap25_2430, Target_Tap25_2440, Target_Tap25_2450, Target_Tap25_2470, Target_Tap25_2480,
                                      Target_Tap25_2490, Target_Tap25_2500, Target_Tap25_2510, Target_Tap25_2520, Target_Tap25_2530, Target_Tap25_2540,
                                      Target_Tap25_2550, Target_Tap25_2560, Target_Tap25_2570, Target_Tap25_2580, Target_Tap25_2590, Target_Tap25_2600,
                                      Target_Tap25_2610, Target_Tap25_2620, Target_Tap25_2640, Target_Tap25_2650, Target_Tap25_2660, Target_Tap25_2680,
                                      Target_Tap25_2690, Target_Tap25_2700, Target_Tap25_2710, Target_Tap25_2720, Target_Tap25_2730, Target_Tap25_2750,
                                      Target_Tap25_2760, Target_Tap25_2770, Target_Tap25_2780, Target_Tap25_2790, Target_Tap25_2800, Target_Tap25_2820,
                                      Target_Tap25_2830, Target_Tap25_2840, Target_Tap25_2850, Target_Tap25_2860, Target_Tap25_2870, Target_Tap25_2890,
                                      Target_Tap25_2900, Target_Tap25_2910, Target_Tap25_2920, Target_Tap25_2940, Target_Tap25_2950, Target_Tap25_2960,
                                      Target_Tap25_2980, Target_Tap25_2990, Target_Tap25_3000, Target_Tap25_3010, Target_Tap25_3020, Target_Tap25_3030,
                                      Target_Tap25_3050, Target_Tap25_3060, Target_Tap25_3070, Target_Tap25_3080, Target_Tap25_3090, Target_Tap25_3100,
                                      Target_Tap25_3120, Target_Tap25_3130, Target_Tap25_3140, Target_Tap25_3150, Target_Tap25_3160, Target_Tap25_3170,
                                      Target_Tap25_3190, Target_Tap25_3200, Target_Tap25_3210, Target_Tap25_3220, Target_Tap25_3230, Target_Tap25_3240,
                                      Target_Tap25_3250, Target_Tap25_3260, Target_Tap25_3270];
        CONST robtarget p_vacio_25{48}:=[Target_Tap25_10, Target_Tap25_80, Target_Tap25_160, Target_Tap25_230, Target_Tap25_330, Target_Tap25_430, Target_Tap25_490,
                                       Target_Tap25_530, Target_Tap25_600, Target_Tap25_680, Target_Tap25_720, Target_Tap25_750, Target_Tap25_820, Target_Tap25_910,
                                       Target_Tap25_1010, Target_Tap25_1070, Target_Tap25_1120, Target_Tap25_1170, Target_Tap25_1220, Target_Tap25_1310, Target_Tap25_1380,
                                       Target_Tap25_1460, Target_Tap25_1520, Target_Tap25_1610, Target_Tap25_1660, Target_Tap25_1740, Target_Tap25_1790, Target_Tap25_1840,
                                       Target_Tap25_1890, Target_Tap25_1960, Target_Tap25_2050, Target_Tap25_2090, Target_Tap25_2130, Target_Tap25_2190, Target_Tap25_2270,
                                       Target_Tap25_2310, Target_Tap25_2380, Target_Tap25_2460, Target_Tap25_2630, Target_Tap25_2670, Target_Tap25_2740, Target_Tap25_2810,
                                       Target_Tap25_2880, Target_Tap25_2930, Target_Tap25_2970, Target_Tap25_3040, Target_Tap25_3110, Target_Tap25_3180];


    PROC Decorar_Meca25(PERS wobjdata WO_Pastel)
        Mover_a_vacio;
        MoveJ Target_Home_10,Vel_Vacio_Rap,Z_Vacio_Rap,Prototipo_JSDaleman\WObj:=wobj0;
        ReiniciarIndices;
        path_contacto_actual:="p_contacto_25";
        path_vacio_actual:="p_vacio_25";
        Path_Tapa_25meca WO_Pastel;
        Mover_en_vacio;
        MoveJ Target_Home_10,Vel_Vacio_Rap,Z_Vacio_Rap,Prototipo_JSDaleman\WObj:=wobj0;
    ENDPROC

    PROC Path_Tapa_25meca(PERS wobjdata WO_Pastel)
        Path_vacio_ejecucion p_vacio_25, 1, WO_Pastel, FALSE;
        Path_contacto_ejecucion p_contacto_25, 1, 6, WO_Pastel, TRUE;
        Path_vacio_ejecucion p_vacio_25, 2, WO_Pastel, FALSE;
        index_vacio_destino:=13;
        Mover_a_contacto;
        TriggL p_contacto_25{7},Vel_Proceso,triggContacto,Z_Proceso,Prototipo_JSDaleman\WObj:=WO_Pastel;
        Mover_en_contacto;
        TriggC p_contacto_25{8},p_contacto_25{9},Vel_Proceso,triggContactoCir,Z_Proceso,Prototipo_JSDaleman\WObj:=WO_Pastel;
        TriggC p_contacto_25{10},p_contacto_25{11},Vel_Proceso,triggContactoCir,Z_Proceso,Prototipo_JSDaleman\WObj:=WO_Pastel;
        TriggL p_contacto_25{12},Vel_Proceso,triggContacto,Z_Proceso,Prototipo_JSDaleman\WObj:=WO_Pastel;
        Mover_a_vacio;
        TriggL p_contacto_25{13},Vel_Acercamiento,triggContacto,Z_Proceso,Prototipo_JSDaleman\WObj:=WO_Pastel;
        Path_vacio_ejecucion p_vacio_25, 3, WO_Pastel, FALSE;
        index_vacio_destino:=19;
        Mover_a_contacto;
        TriggL p_contacto_25{14},Vel_Acercamiento,triggContacto,Z_Acercamiento,Prototipo_JSDaleman\WObj:=WO_Pastel;
        Mover_en_contacto;
        TriggC p_contacto_25{15},p_contacto_25{16},Vel_Proceso,triggContactoCir,Z_Proceso,Prototipo_JSDaleman\WObj:=WO_Pastel;
        TriggC p_contacto_25{17},p_contacto_25{18},Vel_Proceso,triggContactoCir,Z_Proceso,Prototipo_JSDaleman\WObj:=WO_Pastel;
        Mover_a_vacio;
        TriggL p_contacto_25{19},Vel_Acercamiento,triggContacto,Z_Acercamiento,Prototipo_JSDaleman\WObj:=WO_Pastel;
        Path_vacio_ejecucion p_vacio_25, 4, WO_Pastel, FALSE;
        index_vacio_destino:=28;
        Path_contacto_ejecucion p_contacto_25, 20, 22, WO_Pastel, FALSE;
        Mover_en_contacto;
        TriggC p_contacto_25{23},p_contacto_25{24},Vel_Proceso,triggContactoCir,Z_Proceso,Prototipo_JSDaleman\WObj:=WO_Pastel;
        TriggC p_contacto_25{25},p_contacto_25{26},Vel_Proceso,triggContactoCir,Z_Proceso,Prototipo_JSDaleman\WObj:=WO_Pastel;
        TriggL p_contacto_25{27},Vel_Proceso,triggContacto,Z_Proceso,Prototipo_JSDaleman\WObj:=WO_Pastel;
        Mover_a_vacio;
        TriggL p_contacto_25{28},Vel_Acercamiento,triggContacto,Z_Acercamiento,Prototipo_JSDaleman\WObj:=WO_Pastel;
        Path_vacio_ejecucion p_vacio_25, 5, WO_Pastel, FALSE;
        Path_contacto_ejecucion p_contacto_25, 29, 37, WO_Pastel, TRUE;
        Path_vacio_ejecucion p_vacio_25, 6, WO_Pastel, FALSE;
        Path_contacto_ejecucion p_contacto_25, 38, 42, WO_Pastel, TRUE;
        Path_vacio_ejecucion p_vacio_25, 7, WO_Pastel, FALSE;
        Path_contacto_ejecucion p_contacto_25, 43, 45, WO_Pastel, TRUE;
        Path_vacio_ejecucion p_vacio_25, 8, WO_Pastel, FALSE;
        Mover_a_contacto;
        index_vacio_destino:=51;
        TriggL p_contacto_25{46},Vel_Acercamiento,triggContacto,Z_Acercamiento,Prototipo_JSDaleman\WObj:=WO_Pastel;
        Mover_en_contacto;
        TriggC p_contacto_25{47},p_contacto_25{48},Vel_Proceso,triggContactoCir,Z_Proceso,Prototipo_JSDaleman\WObj:=WO_Pastel;
        TriggC p_contacto_25{49},p_contacto_25{50},Vel_Proceso,triggContactoCir,Z_Proceso,Prototipo_JSDaleman\WObj:=WO_Pastel;
        Mover_a_vacio;
        TriggL p_contacto_25{51},Vel_Acercamiento,triggContacto,Z_Acercamiento,Prototipo_JSDaleman\WObj:=WO_Pastel;
        Path_vacio_ejecucion p_vacio_25, 9, WO_Pastel, FALSE;
        Path_contacto_ejecucion p_contacto_25, 52, 58, WO_Pastel, TRUE;
        Path_vacio_ejecucion p_vacio_25, 10, WO_Pastel, FALSE;
        Path_contacto_ejecucion p_contacto_25, 59, 61, WO_Pastel, TRUE;
        Path_vacio_ejecucion p_vacio_25, 11, WO_Pastel, FALSE;
        Path_contacto_ejecucion p_contacto_25, 62, 63, WO_Pastel, TRUE;
        Path_vacio_ejecucion p_vacio_25, 12, WO_Pastel, FALSE;
        index_vacio_destino:=69;
        Mover_a_contacto;
        TriggL p_contacto_25{64},Vel_Acercamiento,triggContacto,Z_Acercamiento,Prototipo_JSDaleman\WObj:=WO_Pastel;
        Mover_en_contacto;
        TriggC p_contacto_25{65},p_contacto_25{66},Vel_Proceso,triggContactoCir,Z_Proceso,Prototipo_JSDaleman\WObj:=WO_Pastel;
        TriggC p_contacto_25{67},p_contacto_25{68},Vel_Proceso,triggContactoCir,Z_Proceso,Prototipo_JSDaleman\WObj:=WO_Pastel;
        Mover_a_vacio;
        TriggL p_contacto_25{69},Vel_Acercamiento,triggContacto,Z_Acercamiento,Prototipo_JSDaleman\WObj:=WO_Pastel;
        Path_vacio_ejecucion p_vacio_25, 13, WO_Pastel, FALSE;
        index_vacio_destino:=77;
        Mover_a_contacto;
        Path_contacto_ejecucion p_contacto_25, 70, 72, WO_Pastel, FALSE;
        Mover_en_contacto;
        TriggC p_contacto_25{73},p_contacto_25{74},Vel_Proceso,triggContactoCir,Z_Proceso,Prototipo_JSDaleman\WObj:=WO_Pastel;
        TriggC p_contacto_25{75},p_contacto_25{76},Vel_Proceso,triggContactoCir,Z_Proceso,Prototipo_JSDaleman\WObj:=WO_Pastel;
        Mover_a_vacio;
        TriggL p_contacto_25{77},Vel_Acercamiento,triggContacto,Z_Acercamiento,Prototipo_JSDaleman\WObj:=WO_Pastel;
        Path_vacio_ejecucion p_vacio_25, 14, WO_Pastel, FALSE;
        index_vacio_destino:=86;
        Mover_a_contacto;
        TriggL p_contacto_25{78},Vel_Acercamiento,triggContacto,Z_Acercamiento,Prototipo_JSDaleman\WObj:=WO_Pastel;
        Mover_en_contacto;
        TriggC p_contacto_25{79},p_contacto_25{80},Vel_Proceso,triggContactoCir,Z_Proceso,Prototipo_JSDaleman\WObj:=WO_Pastel;
        TriggC p_contacto_25{81},p_contacto_25{82},Vel_Proceso,triggContactoCir,Z_Proceso,Prototipo_JSDaleman\WObj:=WO_Pastel;
        TriggL p_contacto_25{83},Vel_Proceso,triggContacto,Z_Proceso,Prototipo_JSDaleman\WObj:=WO_Pastel;
        TriggL p_contacto_25{84},Vel_Proceso,triggContacto,Z_Proceso,Prototipo_JSDaleman\WObj:=WO_Pastel;
        TriggL p_contacto_25{85},Vel_Proceso,triggContacto,Z_Proceso,Prototipo_JSDaleman\WObj:=WO_Pastel;
        Mover_a_vacio;
        TriggL p_contacto_25{86},Vel_Acercamiento,triggContacto,Z_Acercamiento,Prototipo_JSDaleman\WObj:=WO_Pastel;
        Path_vacio_ejecucion p_vacio_25, 15, WO_Pastel, FALSE;
        Path_contacto_ejecucion p_contacto_25, 87, 91, WO_Pastel, TRUE;
        Path_vacio_ejecucion p_vacio_25, 16, WO_Pastel, FALSE;
        index_vacio_destino:=95;
        Mover_a_contacto;
        TriggL p_contacto_25{92},Vel_Acercamiento,triggContacto,Z_Acercamiento,Prototipo_JSDaleman\WObj:=WO_Pastel;
        Mover_en_contacto;
        TriggC p_contacto_25{93},p_contacto_25{94},Vel_Proceso,triggContactoCir,Z_Proceso,Prototipo_JSDaleman\WObj:=WO_Pastel;
        Mover_a_vacio;
        TriggL p_contacto_25{95},Vel_Acercamiento,triggContacto,Z_Acercamiento,Prototipo_JSDaleman\WObj:=WO_Pastel;
        Path_vacio_ejecucion p_vacio_25, 17, WO_Pastel, FALSE;
        index_vacio_destino:=99;
        Mover_a_contacto;
        TriggL p_contacto_25{96},Vel_Acercamiento,triggContacto,Z_Acercamiento,Prototipo_JSDaleman\WObj:=WO_Pastel;
        Mover_en_contacto;
        TriggC p_contacto_25{97},p_contacto_25{98},Vel_Proceso,triggContactoCir,Z_Proceso,Prototipo_JSDaleman\WObj:=WO_Pastel;
        Mover_a_vacio;
        TriggL p_contacto_25{99},Vel_Acercamiento,triggContacto,Z_Acercamiento,Prototipo_JSDaleman\WObj:=WO_Pastel;
        Path_vacio_ejecucion p_vacio_25, 18, WO_Pastel, FALSE;
        index_vacio_destino:=103;
        Mover_a_contacto;
        TriggL p_contacto_25{100},Vel_Acercamiento,triggContacto,Z_Acercamiento,Prototipo_JSDaleman\WObj:=WO_Pastel;
        Mover_en_contacto;
        TriggC p_contacto_25{101},p_contacto_25{102},Vel_Proceso,triggContactoCir,Z_Proceso,Prototipo_JSDaleman\WObj:=WO_Pastel;
        Mover_a_vacio;
        TriggL p_contacto_25{103},Vel_Acercamiento,triggContacto,Z_Acercamiento,Prototipo_JSDaleman\WObj:=WO_Pastel;
        Path_vacio_ejecucion p_vacio_25, 19, WO_Pastel, FALSE;
        index_vacio_destino:=111;
        Mover_a_contacto;
        TriggL p_contacto_25{104},Vel_Acercamiento,triggContacto,Z_Acercamiento,Prototipo_JSDaleman\WObj:=WO_Pastel;
        Mover_en_contacto;
        TriggC p_contacto_25{105},p_contacto_25{106},Vel_Proceso,triggContactoCir,Z_Proceso,Prototipo_JSDaleman\WObj:=WO_Pastel;
        TriggL p_contacto_25{107},Vel_Proceso,triggContacto,Z_Proceso,Prototipo_JSDaleman\WObj:=WO_Pastel;
        TriggL p_contacto_25{108},Vel_Proceso,triggContacto,Z_Proceso,Prototipo_JSDaleman\WObj:=WO_Pastel;
        TriggC p_contacto_25{109},p_contacto_25{110},Vel_Proceso,triggContactoCir,Z_Proceso,Prototipo_JSDaleman\WObj:=WO_Pastel;
        Mover_a_vacio;
        TriggL p_contacto_25{111},Vel_Vacio,triggContacto,Z_VacioMov,Prototipo_JSDaleman\WObj:=WO_Pastel;
        Path_vacio_ejecucion p_vacio_25, 20, WO_Pastel, FALSE;
        index_vacio_destino:=117;
        Mover_a_contacto;
        TriggL p_contacto_25{112},Vel_Acercamiento,triggContacto,Z_Acercamiento,Prototipo_JSDaleman\WObj:=WO_Pastel;
        Mover_en_contacto;
        TriggC p_contacto_25{113},p_contacto_25{114},Vel_Proceso,triggContactoCir,Z_Proceso,Prototipo_JSDaleman\WObj:=WO_Pastel;
        TriggC p_contacto_25{115},p_contacto_25{116},Vel_Proceso,triggContactoCir,Z_Proceso,Prototipo_JSDaleman\WObj:=WO_Pastel;
        Mover_a_vacio;
        TriggL p_contacto_25{117},Vel_Acercamiento,triggContacto,Z_Acercamiento,Prototipo_JSDaleman\WObj:=WO_Pastel;
        Path_vacio_ejecucion p_vacio_25, 21, WO_Pastel, FALSE;
        index_vacio_destino:=124;
        Mover_a_contacto;
        TriggL p_contacto_25{118},Vel_Acercamiento,triggContacto,Z_Acercamiento,Prototipo_JSDaleman\WObj:=WO_Pastel;
        Mover_en_contacto;
        TriggL p_contacto_25{119},Vel_Proceso,triggContacto,Z_Proceso,Prototipo_JSDaleman\WObj:=WO_Pastel;
        TriggC p_contacto_25{120},p_contacto_25{121},Vel_Proceso,triggContactoCir,Z_Proceso,Prototipo_JSDaleman\WObj:=WO_Pastel;
        TriggL p_contacto_25{122},Vel_Proceso,triggContacto,Z_Proceso,Prototipo_JSDaleman\WObj:=WO_Pastel;
        TriggL p_contacto_25{123},Vel_Proceso,triggContacto,Z_Proceso,Prototipo_JSDaleman\WObj:=WO_Pastel;
        Mover_a_vacio;
        TriggL p_contacto_25{124},Vel_Acercamiento,triggContacto,Z_Acercamiento,Prototipo_JSDaleman\WObj:=WO_Pastel;
        Path_vacio_ejecucion p_vacio_25, 22, WO_Pastel, FALSE;
        Path_contacto_ejecucion p_contacto_25, 125, 129, WO_Pastel, TRUE;
        Path_vacio_ejecucion p_vacio_25, 23, WO_Pastel, FALSE;
        index_vacio_destino:=137;
        Path_contacto_ejecucion p_contacto_25, 130, 132, WO_Pastel, FALSE;
        Mover_en_contacto;
        TriggC p_contacto_25{133},p_contacto_25{134},Vel_Proceso,triggContactoCir,Z_Proceso,Prototipo_JSDaleman\WObj:=WO_Pastel;
        TriggC p_contacto_25{135},p_contacto_25{136},Vel_Proceso,triggContactoCir,Z_Proceso,Prototipo_JSDaleman\WObj:=WO_Pastel;
        Mover_a_vacio;
        TriggL p_contacto_25{137},Vel_Acercamiento,triggContacto,Z_Acercamiento,Prototipo_JSDaleman\WObj:=WO_Pastel;
        Path_vacio_ejecucion p_vacio_25, 24, WO_Pastel, FALSE;
        Path_contacto_ejecucion p_contacto_25, 138, 141, WO_Pastel, TRUE;
        Path_vacio_ejecucion p_vacio_25, 25, WO_Pastel, FALSE;
        index_vacio_destino:=148;
        Mover_a_contacto;
        TriggL p_contacto_25{142},Vel_Acercamiento,triggContacto,Z_Acercamiento,Prototipo_JSDaleman\WObj:=WO_Pastel;
        Mover_en_contacto;
        TriggC p_contacto_25{143},p_contacto_25{144},Vel_Proceso,triggContactoCir,Z_Proceso,Prototipo_JSDaleman\WObj:=WO_Pastel;
        TriggC p_contacto_25{145},p_contacto_25{146},Vel_Proceso,triggContactoCir,Z_Proceso,Prototipo_JSDaleman\WObj:=WO_Pastel;
        TriggL p_contacto_25{147},Vel_Proceso,triggContacto,Z_Proceso,Prototipo_JSDaleman\WObj:=WO_Pastel;
        Mover_a_vacio;
        TriggL p_contacto_25{148},Vel_Acercamiento,triggContacto,Z_Acercamiento,Prototipo_JSDaleman\WObj:=WO_Pastel;
        Path_vacio_ejecucion p_vacio_25, 26, WO_Pastel, FALSE;
        index_vacio_destino:=152;
        Mover_a_contacto;
        TriggL p_contacto_25{149},Vel_Acercamiento,triggContacto,Z_Acercamiento,Prototipo_JSDaleman\WObj:=WO_Pastel;
        Mover_en_contacto;
        TriggC p_contacto_25{150},p_contacto_25{151},Vel_Proceso,triggContactoCir,Z_Proceso,Prototipo_JSDaleman\WObj:=WO_Pastel;
        Mover_en_vacio;
        TriggL p_contacto_25{152},Vel_Acercamiento,triggContacto,Z_Acercamiento,Prototipo_JSDaleman\WObj:=WO_Pastel;
        Path_vacio_ejecucion p_vacio_25, 27, WO_Pastel, FALSE;
        index_vacio_destino:=156;
        Mover_a_contacto;
        TriggL p_contacto_25{153},Vel_Acercamiento,triggContacto,Z_Acercamiento,Prototipo_JSDaleman\WObj:=WO_Pastel;
        Mover_en_contacto;
        TriggC p_contacto_25{154},p_contacto_25{155},Vel_Proceso,triggContactoCir,Z_Proceso,Prototipo_JSDaleman\WObj:=WO_Pastel;
        Mover_a_vacio;
        TriggL p_contacto_25{156},Vel_Acercamiento,triggContacto,Z_Acercamiento,Prototipo_JSDaleman\WObj:=WO_Pastel;
        Path_vacio_ejecucion p_vacio_25, 28, WO_Pastel, FALSE;
        Path_contacto_ejecucion p_contacto_25, 157, 160, WO_Pastel, TRUE;
        Path_vacio_ejecucion p_vacio_25, 29, WO_Pastel, FALSE;
        Path_contacto_ejecucion p_contacto_25, 161, 166, WO_Pastel, TRUE;
        Path_vacio_ejecucion p_vacio_25, 30, WO_Pastel, FALSE;
        index_vacio_destino:=174;
        Path_contacto_ejecucion p_contacto_25, 167, 169, WO_Pastel, FALSE;
        Mover_en_contacto;
        TriggC p_contacto_25{170},p_contacto_25{171},Vel_Proceso,triggContactoCir,Z_Proceso,Prototipo_JSDaleman\WObj:=WO_Pastel;
        TriggC p_contacto_25{172},p_contacto_25{173},Vel_Proceso,triggContactoCir,Z_Proceso,Prototipo_JSDaleman\WObj:=WO_Pastel;
        Mover_a_vacio;
        TriggL p_contacto_25{174},Vel_Acercamiento,triggContacto,Z_Acercamiento,Prototipo_JSDaleman\WObj:=WO_Pastel;
        Path_vacio_ejecucion p_vacio_25, 31, WO_Pastel, FALSE;
        Path_contacto_ejecucion p_contacto_25, 175, 177, WO_Pastel, TRUE;
        Path_vacio_ejecucion p_vacio_25, 32, WO_Pastel, FALSE;
        Path_contacto_ejecucion p_contacto_25, 178, 180, WO_Pastel, TRUE;
        Path_vacio_ejecucion p_vacio_25, 33, WO_Pastel, FALSE;
        Path_contacto_ejecucion p_contacto_25, 181, 185, WO_Pastel, TRUE;
        Path_vacio_ejecucion p_vacio_25, 34, WO_Pastel, FALSE;
        index_vacio_destino:=192;
        Mover_a_contacto;
        TriggL p_contacto_25{186},Vel_Acercamiento,triggContacto,Z_Acercamiento,Prototipo_JSDaleman\WObj:=WO_Pastel;
        Mover_en_contacto;
        TriggC p_contacto_25{187},p_contacto_25{188},Vel_Proceso,triggContactoCir,Z_Proceso,Prototipo_JSDaleman\WObj:=WO_Pastel;
        TriggC p_contacto_25{189},p_contacto_25{190},Vel_Proceso,triggContactoCir,Z_Proceso,Prototipo_JSDaleman\WObj:=WO_Pastel;
        TriggL p_contacto_25{191},Vel_Proceso,triggContacto,Z_Proceso,Prototipo_JSDaleman\WObj:=WO_Pastel;
        Mover_a_vacio;
        TriggL p_contacto_25{192},Vel_Acercamiento,triggContacto,Z_Acercamiento,Prototipo_JSDaleman\WObj:=WO_Pastel;
        Path_vacio_ejecucion p_vacio_25, 35, WO_Pastel, FALSE;
        Path_contacto_ejecucion p_contacto_25, 193, 195, WO_Pastel, TRUE;
        Path_vacio_ejecucion p_vacio_25, 36, WO_Pastel, FALSE;
        Path_contacto_ejecucion p_contacto_25, 196, 201, WO_Pastel, TRUE;
        Path_vacio_ejecucion p_vacio_25, 37, WO_Pastel, FALSE;
        index_vacio_destino:=208;
        Mover_a_contacto;
        TriggL p_contacto_25{202},Vel_Acercamiento,triggContacto,Z_Acercamiento,Prototipo_JSDaleman\WObj:=WO_Pastel;
        Mover_en_contacto;
        TriggC p_contacto_25{203},p_contacto_25{204},Vel_Proceso,triggContactoCir,Z_Proceso,Prototipo_JSDaleman\WObj:=WO_Pastel;
        TriggC p_contacto_25{205},p_contacto_25{206},Vel_Proceso,triggContactoCir,Z_Proceso,Prototipo_JSDaleman\WObj:=WO_Pastel;
        TriggL p_contacto_25{207},Vel_Proceso,triggContacto,Z_Proceso,Prototipo_JSDaleman\WObj:=WO_Pastel;
        Mover_a_vacio;
        TriggL p_contacto_25{208},Vel_Acercamiento,triggContacto,Z_Acercamiento,Prototipo_JSDaleman\WObj:=WO_Pastel;
        Path_vacio_ejecucion p_vacio_25, 38, WO_Pastel, FALSE;
        index_vacio_destino:=224;
        Mover_a_contacto;
        TriggL p_contacto_25{209},Vel_Acercamiento,triggContacto,Z_Acercamiento,Prototipo_JSDaleman\WObj:=WO_Pastel;
        Mover_en_contacto;
        TriggC p_contacto_25{210},p_contacto_25{211},Vel_Proceso,triggContactoCir,Z_Proceso,Prototipo_JSDaleman\WObj:=WO_Pastel;
        TriggL p_contacto_25{212},Vel_Proceso,triggContacto,Z_Proceso,Prototipo_JSDaleman\WObj:=WO_Pastel;
        TriggC p_contacto_25{213},p_contacto_25{214},Vel_Proceso,triggContactoCir,Z_Proceso,Prototipo_JSDaleman\WObj:=WO_Pastel;
        TriggC p_contacto_25{215},p_contacto_25{216},Vel_Proceso,triggContactoCir,Z_Proceso,Prototipo_JSDaleman\WObj:=WO_Pastel;
        TriggL p_contacto_25{217},Vel_Acercamiento,triggContacto,Z_Acercamiento,Prototipo_JSDaleman\WObj:=WO_Pastel;
        TriggL p_contacto_25{218},Vel_Proceso,triggContacto,Z_Proceso,Prototipo_JSDaleman\WObj:=WO_Pastel;
        TriggL p_contacto_25{219},Vel_Acercamiento,triggContacto,Z_Acercamiento,Prototipo_JSDaleman\WObj:=WO_Pastel;
        TriggL p_contacto_25{220},Vel_Proceso,triggContacto,Z_Proceso,Prototipo_JSDaleman\WObj:=WO_Pastel;
        TriggL p_contacto_25{221},Vel_Proceso,triggContacto,Z_Proceso,Prototipo_JSDaleman\WObj:=WO_Pastel;
        TriggL p_contacto_25{222},Vel_Proceso,triggContacto,Z_Proceso,Prototipo_JSDaleman\WObj:=WO_Pastel;
        TriggL p_contacto_25{223},Vel_Proceso,triggContacto,Z_Proceso,Prototipo_JSDaleman\WObj:=WO_Pastel;
        Mover_a_vacio;
        TriggL p_contacto_25{224},Vel_Acercamiento,triggContacto,Z_Acercamiento,Prototipo_JSDaleman\WObj:=WO_Pastel;
        Path_vacio_ejecucion p_vacio_25, 39, WO_Pastel, FALSE;
        Path_contacto_ejecucion p_contacto_25, 225, 227, WO_Pastel, TRUE;
        Path_vacio_ejecucion p_vacio_25, 40, WO_Pastel, TRUE;
        index_vacio_destino:=233;
        Mover_a_contacto;
        TriggL p_contacto_25{228},Vel_Acercamiento,triggContacto,Z_Acercamiento,Prototipo_JSDaleman\WObj:=WO_Pastel;
        Mover_en_contacto;
        TriggC p_contacto_25{229},p_contacto_25{230},Vel_Proceso,triggContactoCir,Z_Proceso,Prototipo_JSDaleman\WObj:=WO_Pastel;
        TriggL p_contacto_25{231},Vel_Proceso,triggContacto,Z_Proceso,Prototipo_JSDaleman\WObj:=WO_Pastel;
        TriggL p_contacto_25{232},Vel_Proceso,triggContacto,Z_Proceso,Prototipo_JSDaleman\WObj:=WO_Pastel;
        Mover_a_vacio;
        TriggL p_contacto_25{233},Vel_Acercamiento,triggContacto,Z_Acercamiento,Prototipo_JSDaleman\WObj:=WO_Pastel;
        Path_vacio_ejecucion p_vacio_25, 41, WO_Pastel, FALSE;
        index_vacio_destino:=239;
        Mover_a_contacto;
        TriggL p_contacto_25{234},Vel_Acercamiento,triggContacto,Z_Acercamiento,Prototipo_JSDaleman\WObj:=WO_Pastel;
        Mover_en_contacto;
        TriggC p_contacto_25{235},p_contacto_25{236},Vel_Proceso,triggContactoCir,Z_Proceso,Prototipo_JSDaleman\WObj:=WO_Pastel;
        TriggC p_contacto_25{237},p_contacto_25{238},Vel_Proceso,triggContactoCir,Z_Proceso,Prototipo_JSDaleman\WObj:=WO_Pastel;
        Mover_a_vacio;
        TriggL p_contacto_25{239},Vel_Acercamiento,triggContacto,Z_Acercamiento,Prototipo_JSDaleman\WObj:=WO_Pastel;
        Path_vacio_ejecucion p_vacio_25, 42, WO_Pastel, FALSE;
        index_vacio_destino:=245;
        Mover_a_vacio;
        TriggL p_contacto_25{240},Vel_Acercamiento,triggContacto,Z_Acercamiento,Prototipo_JSDaleman\WObj:=WO_Pastel;
        Mover_en_contacto;
        TriggC p_contacto_25{241},p_contacto_25{242},Vel_Proceso,triggContactoCir,Z_Proceso,Prototipo_JSDaleman\WObj:=WO_Pastel;
        TriggC p_contacto_25{243},p_contacto_25{244},Vel_Proceso,triggContactoCir,Z_Proceso,Prototipo_JSDaleman\WObj:=WO_Pastel;
        Mover_a_vacio;
        TriggL p_contacto_25{245},Vel_Acercamiento,triggContacto,Z_Acercamiento,Prototipo_JSDaleman\WObj:=WO_Pastel;
        Path_vacio_ejecucion p_vacio_25, 43, WO_Pastel, FALSE;
        Path_contacto_ejecucion p_contacto_25, 246, 249, WO_Pastel, TRUE;
        Path_vacio_ejecucion p_vacio_25, 44, WO_Pastel, FALSE;
        Path_contacto_ejecucion p_contacto_25, 250, 252, WO_Pastel, TRUE;
        Path_vacio_ejecucion p_vacio_25, 45, WO_Pastel, FALSE;
        index_vacio_destino:=258;
        Mover_a_contacto;
        TriggL p_contacto_25{253},Vel_Acercamiento,triggContacto,Z_Acercamiento,Prototipo_JSDaleman\WObj:=WO_Pastel;
        Mover_en_contacto;
        TriggC p_contacto_25{254},p_contacto_25{255},Vel_Proceso,triggContactoCir,Z_Proceso,Prototipo_JSDaleman\WObj:=WO_Pastel;
        TriggL p_contacto_25{256},Vel_Proceso,triggContacto,Z_Proceso,Prototipo_JSDaleman\WObj:=WO_Pastel;
        TriggL p_contacto_25{257},Vel_Proceso,triggContacto,Z_Proceso,Prototipo_JSDaleman\WObj:=WO_Pastel;
        Mover_a_vacio;
        TriggL p_contacto_25{258},Vel_Acercamiento,triggContacto,Z_Acercamiento,Prototipo_JSDaleman\WObj:=WO_Pastel;
        Path_vacio_ejecucion p_vacio_25, 46, WO_Pastel, FALSE;
        index_vacio_destino:=264;
        Mover_a_contacto;
        TriggL p_contacto_25{259},Vel_Acercamiento,triggContacto,Z_Acercamiento,Prototipo_JSDaleman\WObj:=WO_Pastel;
        Mover_en_contacto;
        TriggC p_contacto_25{260},p_contacto_25{261},Vel_Proceso,triggContactoCir,Z_Proceso,Prototipo_JSDaleman\WObj:=WO_Pastel;
        TriggC p_contacto_25{262},p_contacto_25{263},Vel_Proceso,triggContactoCir,Z_Proceso,Prototipo_JSDaleman\WObj:=WO_Pastel;
        Mover_a_vacio;
        TriggL p_contacto_25{264},Vel_Acercamiento,triggContacto,Z_Acercamiento,Prototipo_JSDaleman\WObj:=WO_Pastel;
        Path_vacio_ejecucion p_vacio_25, 47, WO_Pastel, FALSE;
        index_vacio_destino:=270;
        Mover_a_contacto;
        TriggL p_contacto_25{265},Vel_Acercamiento,triggContacto,Z_Acercamiento,Prototipo_JSDaleman\WObj:=WO_Pastel;
        Mover_en_contacto;
        TriggC p_contacto_25{266},p_contacto_25{267},Vel_Proceso,triggContactoCir,Z_Proceso,Prototipo_JSDaleman\WObj:=WO_Pastel;
        TriggL p_contacto_25{268},Vel_Proceso,triggContacto,Z_Proceso,Prototipo_JSDaleman\WObj:=WO_Pastel;
        TriggL p_contacto_25{269},Vel_Proceso,triggContacto,Z_Proceso,Prototipo_JSDaleman\WObj:=WO_Pastel;
        Mover_a_vacio;
        TriggL p_contacto_25{270},Vel_Acercamiento,triggContacto,Z_Acercamiento,Prototipo_JSDaleman\WObj:=WO_Pastel;
        Path_vacio_ejecucion p_vacio_25, 48, WO_Pastel, FALSE;
        index_vacio_destino:=279;
        Mover_a_contacto;
        TriggL p_contacto_25{271},Vel_Acercamiento,triggContacto,Z_Acercamiento,Prototipo_JSDaleman\WObj:=WO_Pastel;
        Mover_en_contacto;
        TriggC p_contacto_25{272},p_contacto_25{273},Vel_Proceso,triggContactoCir,Z_Proceso,Prototipo_JSDaleman\WObj:=WO_Pastel;
        TriggC p_contacto_25{274},p_contacto_25{275},Vel_Proceso,triggContactoCir,Z_Proceso,Prototipo_JSDaleman\WObj:=WO_Pastel;
        TriggC p_contacto_25{276},p_contacto_25{277},Vel_Proceso,triggContactoCir,Z_Proceso,Prototipo_JSDaleman\WObj:=WO_Pastel;
        TriggL p_contacto_25{278},Vel_Proceso,triggContacto,Z_Proceso,Prototipo_JSDaleman\WObj:=WO_Pastel;
        Mover_a_vacio;
        TriggL p_contacto_25{279},Vel_Acercamiento,triggContacto,Z_Acercamiento,Prototipo_JSDaleman\WObj:=WO_Pastel;
    ENDPROC
ENDMODULE

--- Controller Data/IRB140_LabSIR/RAPID/TASK1/PROGMOD/ModuloPrin.mod ---
MODULE ModuloPrin
    !***********************************************************
    !
    ! Modulo:  ModuloPrin
    !
    ! Descripci?n:
    !   Modulo de inicio para el programa con:
    !   - main: Inicio de la rutina,
    !     inicializaci?n de varibles e interrupciones y proceso principal
    !   - Path_Home_Run: Rutina para llegar al punto de Home del robot
    !   - Path_Transicion: Rutina para punto que evita problemas de mecanismo en home
    !     y transici?n entre rutinas o puntos importantes
    !
    ! Autor: Juan_Daleman
    !
    ! Versi?n: 1.0
    !
    !***********************************************************

    !Puntos de espera y mantenimiento
    CONST robtarget Target_Mantenimiento:=[[524.308309139,712.143242458,575.732],[0.472131723,-0.518247718,0.524360327,-0.483277546],[0,0,0,0],[9E+09,9E+09,9E+09,9E+09,9E+09,9E+09]];
    CONST robtarget Target_Espera:=[[0,-407.163,1030.849],[0.5,0.5,0.5,-0.5],[0,0,0,0],[9E+09,9E+09,9E+09,9E+09,9E+09,9E+09]];

    !Puntos para Home
    !CONST robtarget Target_Home_10:=[[802.284,0,778.685],[0.382683432,0,0.923879533,0],[0,0,0,0],[9E+09,9E+09,9E+09,9E+09,9E+09,9E+09]];
    CONST robtarget Target_Home_10:=[[329.136851055,0,730.080138956],[0.26115172,0,0.965297767,0],[0,0,0,0],[9E+09,9E+09,9E+09,9E+09,9E+09,9E+09]];
    CONST robtarget Target_Home_20:=[[788.429,0,593.609],[0.382683432,0,0.923879533,0],[0,0,0,0],[9E+09,9E+09,9E+09,9E+09,9E+09,9E+09]];

